(* CODESYS project Intecre_TwinSafeModels.library
   Author: Mark Lazarides
   Version: 0.5.0.3
   Description: Functional models of the TwinSAFE logic function blocks and TwinSAFE group, for trialling safety applications and their interaction with the standard PLC.
      
      0.4.2.0 - T_SafeFunctionBlockBase sets State to Run / Stop before Process; user FBs need no State logic.
      0.4.1.0 - corrects call issue with Example_UserFBs
      
      0.4.0.0 - Adds the eight channel (EL1918) and two channel (EL2912) terminal models.
      0.3.0.0 - Adds User FB examples, demonstrating extension.
   Title: Intecre.TwinSAFE.Models
   DefaultNamespace: Intecre.TwinSAFE.Models
   Placeholder: Intecre.TwinSAFE.Models
   Company: Intecre Ltd

Project tree, tasks and I/O mapping:
  libraries: Intecre.Utilities, * (Intecre Ltd); Tc2_Standard, * (Beckhoff Automation GmbH); Tc2_System, * (Beckhoff Automation GmbH); Tc3_Module, * (Beckhoff Automation GmbH); TcUnit, * (www.tcunit.org)
  Core/
    function F_NormaliseSafeInput [ST]
    function F_SafeInputValue [ST]
    function F_SafeResetTimeOk [ST]
    function block T_SafeConnection [ST]: FB_init, RunStateMachine, SetGroupReference, StateChanged
    function block T_SafeFunctionBlockBase [ST]: ClearDiagBit, ConfigurationOk, FB_init, Process, ReportRefusedConfiguration, SetDiagBit, SetGroupReference
    function block T_SafeGroup [ST]: ConnectionCount, FunctionBlockCount, GroupState, RaiseOnRefusedConfiguration, RegisterConnection, RegisterFunctionBlock, ScanMembers, StateChanged
    function block T_SafeInputPair [ST]
    function block T_SafeInputTerminal [ST]
    function block T_SafeInputTerminal8 [ST]
    function block T_SafeOutputTerminal [ST]
    function block T_SafeOutputTerminal2 [ST]
  DUTs/
    data type E_SafeConnectionError
    data type E_SafeConnectionState
    data type E_SafeEdmState
    data type E_SafeFbState
    data type E_SafeGroupDiag
    data type E_SafeGroupState
    data type E_SafeLatchState
    data type E_SafeMonState
    data type E_SafeMutingState
    data type E_SafeTonState
    data type E_SafeTwoHandState
    data type ST_SafeConnShutdownParameters
    data type ST_SafeEdmParameters
    data type ST_SafeEStopParameters
    data type ST_SafeLatchParameters
    data type ST_SafeLogicParameters
    data type ST_SafeMonParameters
    data type ST_SafeMutingParameters
    data type ST_SafeOpModeParameters
    data type ST_SafeTimerParameters
    data type ST_SafeTwoHandParameters
  Examples/
    Example_UserFbs/
      function block T_SafePulse_UserFB [CFC]: FB_init, Process
      function block T_SafeRTrig_UserFB [CFC]: FB_init, Process
    program PRG_EStopExample [ST]
    program PRG_EStopExample_CFC [CFC]
  FunctionBlocks/
    function block T_SafeAnd [ST]: ConfigurationOk, Process
    function block T_SafeConnShutdown [ST]: ConnShutdownState, FB_init, Process, StateChanged, UpdateDiscrepancyDiag
    function block T_SafeDecouple [ST]: Process
    function block T_SafeEdm [ST]: ConfigurationOk, Process, StateChanged
    function block T_SafeEStop [ST]: ConfigurationOk, EdmInputsOk, EdmInputsTrue, EdmResetOk, EStopState, Process, SetOutputsSafe, StartEdmResetMonitoring, StateChanged, UpdateDiscrepancyDiag
    function block T_SafeMon [ST]: ConfigurationOk, EdmInputsOk, EdmInputsTrue, EdmResetOk, MonState, Process, SetOutputsSafe, StartEdmResetMonitoring, StateChanged, UpdateDiscrepancyDiag
    function block T_SafeMuting [ST]: Actual, AddEvent, Advance, AnySensor, BuildSequence, ConfigurationOk, EdmInputsOk, EdmInputsTrue, EdmResetOk, IsMuting, MutingState, MutingStateFor, Process, SetOutputsSafe, StartEdmResetMonitoring, StateChanged, UpdateDiscrepancyDiag
    function block T_SafeOpMode [ST]: ConfigurationOk, Process, SetOutputs, StateChanged
    function block T_SafeOr [ST]: ConfigurationOk, Process
    function block T_SafeRs [ST]: ConfigurationOk, Process
    function block T_SafeSr [ST]: ConfigurationOk, Process
    function block T_SafeTof [ST]: ConfigurationOk, Process
    function block T_SafeTon [ST]: ConfigurationOk, Process
    function block T_SafeTwoHand [ST]: Process, SetHandDiscrepancyError, StateChanged, TwoHandState, UpdateDiscrepancyDiag
    function block T_SafeXor [ST]: Process
  Params/
    global variables SafeModelParams
  Project Information/
    function F_GetCompany [ST]
    function F_GetTitle [ST]
    function F_GetVersion [ST]
  Tests/
    User_FB_Tests/
      function block T_SafePulse_UserFB_Tests [ST]: Test_InnerBlocksJoinTheGroup, Test_PulseEndsWhenInputDrops, Test_PulseForDelayTimeWhileInputHeld, Test_StoppedGivesNoOutput
      function block T_SafePulse_UserFB_Tests_CFC [ST]: Test_InnerBlocksJoinTheGroup, Test_PulseEndsWhenInputDrops, Test_PulseForDelayTimeWhileInputHeld, Test_StoppedGivesNoOutput
      function block T_SafeRTrig_UserFB_Tests [ST]: Test_InnerBlocksJoinTheGroup, Test_StoppedGivesNoOutput, Test_TriggerForOneCycleOnRisingEdge
      function block T_SafeRTrig_UserFB_Tests_CFC [ST]: Test_InnerBlocksJoinTheGroup, Test_StoppedGivesNoOutput, Test_TriggerForOneCycleOnRisingEdge
    program PRG_TestRunner [ST]
    function block T_SafeAnd_Tests [ST]: Test_AllConnectedInputsTrueGivesRun, Test_OneConnectedInputIsRefused, Test_OneInputFalseGivesSafe, Test_RaiseOnRefusedConfigurationStopsHard, Test_StoppedGivesNoOutput, Test_UnconnectedInputsIgnoredAndMakeContactNegated
    function block T_SafeAnd_Tests_CFC [ST]: Test_AllConnectedInputsTrueGivesRun, Test_OneInputFalseGivesSafe, Test_StoppedGivesNoOutput, Test_UnconnectedInputsIgnoredAndMakeContactNegated
    function block T_SafeCfcTestSuite [ST]: FinishTest, StartTest
    function block T_SafeConnection_Tests [ST]: Test_ComErrorClearedByAcknowledge, Test_StartsUpToDataWhenGroupRuns
    function block T_SafeConnection_Tests_CFC [ST]: Test_ComErrorClearedByAcknowledge, Test_StartsUpToDataWhenGroupRuns
    function block T_SafeConnShutdown_Tests [ST]: Test_DeactivateShutsDownConnection
    function block T_SafeConnShutdown_Tests_CFC [ST]: Test_DeactivateShutsDownConnection
    function block T_SafeDecouple_Tests [ST]: Test_InputsLoopedToOutputsOnlyWhenRunning
    function block T_SafeDecouple_Tests_CFC [ST]: Test_InputsLoopedToOutputsOnlyWhenRunning
    function block T_SafeEdm_Tests [ST]: Test_NoErrorWhenFeedbackFollows, Test_SwitchOnTimeoutGivesError, Test_UnconnectedMon2IsRefused
    function block T_SafeEdm_Tests_CFC [ST]: Test_NoErrorWhenFeedbackFollows, Test_SwitchOnTimeoutGivesError
    function block T_SafeEStop_Tests [ST]: Test_DelayedOutput, Test_DiscrepancyErrorNeedsSafeInputsBeforeAck, Test_EdmErrorAtRestartAndAcknowledge, Test_EStopRequestSwitchesOutputsOffAndBlocksRestart, Test_MakeContactInputRequestsSafeStateOnOne, Test_OutputsOffWhenStopped, Test_ResetTimeOverSixtySecondsIsRefused, Test_RestartHeldBeforeEStopGivesEdmError, Test_StartupRequiresRestartSequence
    function block T_SafeEStop_Tests_CFC [ST]: Test_DelayedOutput, Test_DiscrepancyErrorNeedsSafeInputsBeforeAck, Test_EdmErrorAtRestartAndAcknowledge, Test_EStopRequestSwitchesOutputsOffAndBlocksRestart, Test_MakeContactInputRequestsSafeStateOnOne, Test_OutputsOffWhenStopped, Test_RestartHeldBeforeEStopGivesEdmError, Test_StartupRequiresRestartSequence
    function block T_SafeGroup_Tests [ST]: Test_ConnectionStartupAndComError, Test_FbErrorStopsGroupAndErrAckRecovers, Test_RefusesTheSixtyFifthConnection, Test_RegistersMoreThanSixtyFourBlocks, Test_RunsFunctionBlocksWithoutConnections, Test_StopWhenRunFalse
    function block T_SafeGroup_Tests_CFC [ST]: Test_ConnectionStartupAndComError, Test_FbErrorStopsGroupAndErrAckRecovers, Test_RunsFunctionBlocksWithoutConnections, Test_StopWhenRunFalse
    function block T_SafeInputPair_Tests [ST]: Test_BreakContactRequestsSafeStateOnZero, Test_DiscrepancyErrorAfterTimeoutAndResetAfterSafeInputs, Test_InactivePairNeverRequestsSafeState, Test_MakeContactRequestsSafeStateOnOne, Test_TwoChannelRequestsSafeStateIfEitherChannelLow
    function block T_SafeInputPair_Tests_CFC [ST]: Test_BreakContactRequestsSafeStateOnZero, Test_DiscrepancyErrorAfterTimeoutAndResetAfterSafeInputs, Test_InactivePairNeverRequestsSafeState, Test_MakeContactRequestsSafeStateOnOne, Test_TwoChannelRequestsSafeStateIfEitherChannelLow
    function block T_SafeInputTerminal8_Tests [ST]: Test_ComErrorForcesSafeInputsFalse, Test_RegistersAsConnection, Test_SafeInputsFalseBeforeData, Test_SafeInputsFollowChannelsInData
    function block T_SafeMon_Tests [ST]: Test_AutomaticRestartWhenGuardClosed, Test_EdmFaultWithoutManualRestartStaysSafe, Test_ManualFunctionTestRequiresGuardOpenedOnce, Test_NoMonInConnectedIsRefused, Test_ResetTimeNotMultipleOfTenIsRefused, Test_SecureInputBypassesGuard
    function block T_SafeMon_Tests_CFC [ST]: Test_AutomaticRestartWhenGuardClosed, Test_EdmFaultWithoutManualRestartStaysSafe, Test_ManualFunctionTestRequiresGuardOpenedOnce, Test_SecureInputBypassesGuard
    function block T_SafeMuting_Tests [ST]: Test_OssdBlockedWithoutMutingGivesSafe, Test_ResetTimeNotMultipleOfTenIsRefused, Test_SequenceViolationGivesError, Test_SequentialMutingKeepsOutputOn, Test_TwoSensorParallelSequence
    function block T_SafeMuting_Tests_CFC [ST]: Test_OssdBlockedWithoutMutingGivesSafe, Test_SequenceViolationGivesError, Test_SequentialMutingKeepsOutputOn, Test_TwoSensorParallelSequence
    function block T_SafeOpMode_Tests [ST]: Test_ConnectedRestartRequiresRestartSequence, Test_ExactlyOneInputSelectsOutput, Test_OneConnectedInputIsRefused, Test_SlowModeChangeGivesDiscrepancyError
    function block T_SafeOpMode_Tests_CFC [ST]: Test_ConnectedRestartRequiresRestartSequence, Test_ExactlyOneInputSelectsOutput, Test_SlowModeChangeGivesDiscrepancyError
    function block T_SafeOr_Tests [ST]: Test_AllFalseGivesSafe, Test_AnyConnectedInputTrueGivesRun, Test_OneConnectedInputIsRefused
    function block T_SafeOr_Tests_CFC [ST]: Test_AllFalseGivesSafe, Test_AnyConnectedInputTrueGivesRun
    function block T_SafeOutputTerminal2_Tests [ST]: Test_ChannelsFalseBeforeData, Test_ChannelsFollowSafeOutsInData, Test_ComErrorForcesChannelsFalse, Test_GroupNotRunningForcesChannelsFalse, Test_RegistersAsConnection
    function block T_SafeRs_Tests [ST]: Test_ResetDominantLatch, Test_UnconnectedSetIsRefused
    function block T_SafeRs_Tests_CFC [ST]: Test_ResetDominantLatch
    function block T_SafeSr_Tests [ST]: Test_SetDominantLatch, Test_UnconnectedResetIsRefused
    function block T_SafeSr_Tests_CFC [ST]: Test_SetDominantLatch
    function block T_SafeTof_Tests [ST]: Test_OutputDelayedOff, Test_UnconnectedInputIsRefused
    function block T_SafeTof_Tests_CFC [ST]: Test_OutputDelayedOff
    function block T_SafeTon_Tests [ST]: Test_OutputDelayedOn, Test_UnconnectedInputIsRefused
    function block T_SafeTon_Tests_CFC [ST]: Test_OutputDelayedOn
    function block T_SafeTwoHand_Tests [ST]: Test_BothHandsGiveOutputAndReleaseNeedsBothOff, Test_HandDiscrepancyTimeout, Test_SecondHandWithoutFirstGivesTwoHandError
    function block T_SafeTwoHand_Tests_CFC [ST]: Test_BothHandsGiveOutputAndReleaseNeedsBothOff, Test_HandDiscrepancyTimeout, Test_SecondHandWithoutFirstGivesTwoHandError
    function block T_SafeXor_Tests [ST]: Test_ConnectedPairsAreExclusiveOr
    function block T_SafeXor_Tests_CFC [ST]: Test_ConnectedPairsAreExclusiveOr
  Version/
    global variables Global_Version
*)

// DUTs/E_SafeConnectionError
// TwinSAFE connection error codes (low nibble of the connection Diag byte).
{attribute 'qualified_only'}
{attribute 'to_string'}
TYPE
E_SafeConnectionError :
(
    NoError := 0,
    InvalidCommand := 1,
    UnknownCommand := 2,
    InvalidConnectionId := 3,
    InvalidCrc := 4,
    WatchdogElapsed := 5,
    InvalidFsoeAddress := 6,
    InvalidData := 7,
    InvalidComParameterLength := 8,
    InvalidComParameters := 9,
    InvalidUserParameterLength := 10,
    InvalidUserParameters := 11,
    FsoeMasterReset := 12,
    SlaveModuleError := 13,
    OutputModuleError := 14,
    SlaveNotStarted := 15
) BYTE;
END_TYPE

// DUTs/E_SafeConnectionState
// TwinSAFE (FSoE) connection state codes.
{attribute 'qualified_only'}
{attribute 'to_string'}
TYPE
E_SafeConnectionState :
(
    Reset := 100,
    Session := 101,
    Connection := 102,
    Parameter := 103,
    Data := 104,
    Shutdown := 105,
    ShutdownDeactive := 106
) BYTE;
END_TYPE

// DUTs/E_SafeEdmState
// FB EDM state codes.
{attribute 'qualified_only'}
{attribute 'to_string'}
TYPE
E_SafeEdmState :
(
    Undefined := 0,
    Stop := 2,
    Error := 4,
    Reset := 5,
    MonOff := 14,
    MonOn := 15
) BYTE;
END_TYPE

// DUTs/E_SafeFbState
// TwinSAFE function block state codes shared by most FBs (Map State value).
// Error is also the state of a block whose configuration the TwinSAFE Safety Editor refuses (too few
// inputs connected, a required input unwired, an invalid EDM reset time): the block then sets Error,
// diagnostic bit 15 (16#8000), which no TwinSAFE FB uses, and stays in Error through every ErrAck.
// See T_SafeFunctionBlockBase.
{attribute 'qualified_only'}
{attribute 'to_string'}
TYPE
E_SafeFbState :
(
    Undefined := 0,
    Run := 1,
    Stop := 2,
    Safe := 3,
    Error := 4,
    Reset := 5,
    Start := 6,
    ErrorDelay := 7,
    DelayOut := 8
) BYTE;
END_TYPE

// DUTs/E_SafeGroupDiag
// TwinSAFE group diagnostic codes (EL/EJ6910).
{attribute 'qualified_only'}
{attribute 'to_string'}
TYPE
E_SafeGroupDiag :
(
    NoError := 0,
    FbError := 1,
    ComError := 2,
    ModuleError := 3,
    CmpError := 4,
    DeactivateError := 5,
    RestartError := 6
) BYTE;
END_TYPE

// DUTs/E_SafeGroupState
// TwinSAFE group state codes (EL/EJ6910).
{attribute 'qualified_only'}
{attribute 'to_string'}
TYPE
E_SafeGroupState :
(
    Undefined := 0,
    Run := 1,
    Stop := 2,
    Safe := 3,
    Error := 4,
    Reset := 5,
    Start := 6,
    StopError := 7,
    Deactive := 16,
    WaitComError := 17
) BYTE;
END_TYPE

// DUTs/E_SafeLatchState
// FB RS and FB SR state codes.
{attribute 'qualified_only'}
{attribute 'to_string'}
TYPE
E_SafeLatchState :
(
    Undefined := 0,
    Stop := 2,
    Safe := 3,
    Set := 9
) BYTE;
END_TYPE

// DUTs/E_SafeMonState
// FB MON state codes.
{attribute 'qualified_only'}
{attribute 'to_string'}
TYPE
E_SafeMonState :
(
    Undefined := 0,
    Run := 1,
    Stop := 2,
    Safe := 3,
    Error := 4,
    Reset := 5,
    Start := 6,
    ErrorDelay := 7,
    DelayOut := 8,
    FuncTest := 9
) BYTE;
END_TYPE

// DUTs/E_SafeMutingState
// FB MUTING state codes.
{attribute 'qualified_only'}
{attribute 'to_string'}
TYPE
E_SafeMutingState :
(
    Undefined := 0,
    Run := 1,
    Stop := 2,
    Safe := 3,
    Error := 4,
    Reset := 5,
    DelayOut := 8,
    Muting1 := 9,
    Muting2 := 10,
    Muting3 := 11,
    Muting4 := 12,
    Muting5 := 13,
    Muting6 := 14,
    Muting7 := 15,
    Muting8 := 16,
    Muting9 := 17
) BYTE;
END_TYPE

// DUTs/E_SafeTonState
// FB TON state codes.
{attribute 'qualified_only'}
{attribute 'to_string'}
TYPE
E_SafeTonState :
(
    Undefined := 0,
    Run := 1,
    Stop := 2,
    Safe := 3,
    DelayIn := 9
) BYTE;
END_TYPE

// DUTs/E_SafeTwoHandState
// FB TWOHAND state codes.
{attribute 'qualified_only'}
{attribute 'to_string'}
TYPE
E_SafeTwoHandState :
(
    Undefined := 0,
    Run := 1,
    Stop := 2,
    Safe := 3,
    Error := 4,
    Reset := 5,
    OneButton := 11,
    TwoButton := 12,
    Release := 13
) BYTE;
END_TYPE

// DUTs/ST_SafeConnShutdownParameters
// Parameters of FB CONNECTION SHUTDOWN.
TYPE
ST_SafeConnShutdownParameters :
STRUCT
    Deactivate1MakeContact : BOOL;
    Deactivate2MakeContact : BOOL;
    DiscrepancyTime : TIME;
    SafeInputsAfterDiscError : BOOL; // Safety Editor checkbox 'Safe Inputs after Disc Error', FALSE for a new block:
        // TRUE makes both channels of the pair that raised a discrepancy error return to the safe state together
        // before ErrAck can clear it
END_STRUCT
END_TYPE

// DUTs/ST_SafeEdmParameters
// Parameters of FB EDM.
TYPE
ST_SafeEdmParameters :
STRUCT
    Mon1MakeContact : BOOL;
    Mon2MakeContact : BOOL;
    SwitchOnTime : TIME; // Mon2 must become FALSE within this time of Mon1 rising. T#0S disables
    SwitchOffTime : TIME; // Mon2 must become TRUE within this time of Mon1 falling. T#0S disables
END_STRUCT
END_TYPE

// DUTs/ST_SafeEStopParameters
// Parameters of FB ESTOP (port and FB properties of the Safety Editor).
// Ports are active when connected; a pair is two channel when both ports are connected.
TYPE
ST_SafeEStopParameters :
STRUCT
    EStopIn1MakeContact : BOOL; // FALSE = break contact (0 requests the safe state); TRUE = make contact
    EStopIn2MakeContact : BOOL;
    EStopIn3MakeContact : BOOL;
    EStopIn4MakeContact : BOOL;
    EStopIn5MakeContact : BOOL;
    EStopIn6MakeContact : BOOL;
    EStopIn7MakeContact : BOOL;
    EStopIn8MakeContact : BOOL;
    DiscrepancyTime1 : TIME; // EStopIn1 / EStopIn2. T#0S = no discrepancy monitoring
    DiscrepancyTime2 : TIME; // EStopIn3 / EStopIn4
    DiscrepancyTime3 : TIME; // EStopIn5 / EStopIn6
    DiscrepancyTime4 : TIME; // EStopIn7 / EStopIn8
    DelayTime : TIME; // switch-off delay of EStopDelOut
    Edm1ResetTime : TIME; // EL6910: EDM1 must drop within this time of EStopOut switching on. T#0S disables
    Edm2ResetTime : TIME;
    SafeInputsAfterDiscError : BOOL; // Safety Editor checkbox, FALSE for a new block; the EL6910 always applies
        // 'Safe Inputs after Disc Error' to ESTOP whatever the box says (only the EL6900 honours it, and the editor
        // warns when it is TRUE under an EL6910), so the model ignores this value and always behaves as TRUE
END_STRUCT
END_TYPE

// DUTs/ST_SafeLatchParameters
// Parameters of FB RS and FB SR.
TYPE
ST_SafeLatchParameters :
STRUCT
    SetMakeContact : BOOL;
    ResetMakeContact : BOOL;
END_STRUCT
END_TYPE

// DUTs/ST_SafeLogicParameters
// Parameters of FB AND and FB OR. Inputs are active when connected.
TYPE
ST_SafeLogicParameters :
STRUCT
    In1MakeContact : BOOL; // TRUE = the input is negated before the logic operation
    In2MakeContact : BOOL;
    In3MakeContact : BOOL;
    In4MakeContact : BOOL;
    In5MakeContact : BOOL;
    In6MakeContact : BOOL;
    In7MakeContact : BOOL;
    In8MakeContact : BOOL;
END_STRUCT
END_TYPE

// DUTs/ST_SafeMonParameters
// Parameters of FB MON. Manual restart is active when the Restart port is connected.
TYPE
ST_SafeMonParameters :
STRUCT
    MonIn1MakeContact : BOOL;
    MonIn2MakeContact : BOOL;
    MonIn3MakeContact : BOOL;
    MonIn4MakeContact : BOOL;
    Secure1MakeContact : BOOL;
    Secure2MakeContact : BOOL;
    DiscrepancyTime1 : TIME; // MonIn1 / MonIn2
    DiscrepancyTime2 : TIME; // MonIn3 / MonIn4
    SecureDiscrepancyTime : TIME; // Secure1 / Secure2
    DelayTime : TIME; // switch-off delay of MonDelOut
    Edm1ResetTime : TIME;
    Edm2ResetTime : TIME;
    ManualFunctionTest : BOOL; // every connected MonIn pair must request the safe state once after start
    SafeInputsAfterDiscError : BOOL; // Safety Editor checkbox 'Safe Inputs after Disc Error', FALSE for a new block:
        // TRUE makes both channels of the pair that raised a discrepancy error return to the safe state together
        // before ErrAck can clear it
END_STRUCT
END_TYPE

// DUTs/ST_SafeMutingParameters
// Parameters of FB MUTING.
TYPE
ST_SafeMutingParameters :
STRUCT
    SequentialInputs : BOOL; // TRUE: single-channel muting sensors in sequence; FALSE: two two-channel sensors
    MutingIn1MakeContact : BOOL;
    MutingIn2MakeContact : BOOL;
    MutingIn3MakeContact : BOOL;
    MutingIn4MakeContact : BOOL;
    OSSDIn1MakeContact : BOOL;
    OSSDIn2MakeContact : BOOL;
    MutingDiscrepancyTime1 : TIME; // MutingIn1 / MutingIn2 (parallel mode)
    MutingDiscrepancyTime2 : TIME; // MutingIn3 / MutingIn4 (parallel mode)
    OssdDiscrepancyTime : TIME; // OSSDIn1 / OSSDIn2
    FilterTime : TIME; // debounce of the muting inputs (max 500 ms)
    MaxMutingTime : TIME; // max duration of a muting sequence (max 10 min). T#0S disables
    DelayTime : TIME; // switch-off delay of MuteDelOut (max 30 s)
    Edm1ResetTime : TIME;
    Edm2ResetTime : TIME;
    BackwardsMode : BOOL; // EL6910: sequence may also run from the last sensor to the first
    OssdCheckOptional : BOOL; // EL6910: protective device is not part of the sequence check
    SafeInputsAfterDiscError : BOOL; // Safety Editor checkbox 'Safe Inputs after Disc Error', FALSE for a new block:
        // TRUE makes both channels of the pair that raised a discrepancy error return to the safe state together
        // before ErrAck can clear it
END_STRUCT
END_TYPE

// DUTs/ST_SafeOpModeParameters
// Parameters of FB OPMODE. Manual restart is active when the Restart port is connected.
TYPE
ST_SafeOpModeParameters :
STRUCT
    DiscrepancyTime : TIME; // max time during a mode change with none or several inputs set. T#0S disables
END_STRUCT
END_TYPE

// DUTs/ST_SafeTimerParameters
// Parameters of FB TON and FB TOF.
TYPE
ST_SafeTimerParameters :
STRUCT
    MakeContact : BOOL;
    DelayTime : TIME;
END_STRUCT
END_TYPE

// DUTs/ST_SafeTwoHandParameters
// Parameters of FB TWOHAND.
TYPE
ST_SafeTwoHandParameters :
STRUCT
    Twohand1MakeContact : BOOL;
    Twohand2MakeContact : BOOL;
    Twohand3MakeContact : BOOL;
    Twohand4MakeContact : BOOL;
    DiscrepancyTime1 : TIME; // Twohand1 / Twohand2
    DiscrepancyTime2 : TIME; // Twohand3 / Twohand4
    HandDiscrepancyTime : TIME; // max time between actuation of the two hands (max 2500 ms). T#0S disables
    SafeInputsAfterDiscError : BOOL; // Safety Editor checkbox 'Safe Inputs after Disc Error', FALSE for a new block:
        // TRUE makes both channels of the pair that raised a discrepancy error return to the safe state together
        // before ErrAck can clear it
END_STRUCT
END_TYPE

// Params/SafeModelParams
// Library parameters of Intecre.TwinSAFE.Models: the project-wide defaults, set per project in the
// Library Manager's parameter view without rebuilding the library. A parameter list must be constant,
// so the run-time switch lives on T_SafeGroup (RaiseOnRefusedConfiguration), initialised from here.
{attribute 'qualified_only'}
VAR_GLOBAL CONSTANT
    // Default of T_SafeGroup.RaiseOnRefusedConfiguration for every group. TRUE: a block of the group whose
    // configuration the TwinSAFE Safety Editor refuses (see T_SafeFunctionBlockBase) raises
    // RTSEXCPT_IO_CONFIG_ERROR with F_RaiseException after it has reported Error, so the controller stops
    // on the first cycle unless the call is in a __TRY block. FALSE: the block only reports Error,
    // State = Error and diagnostic bit 15, and logs the fault once.
    RAISE_ON_REFUSED_CONFIGURATION : BOOL := FALSE;
END_VAR

// Version/Global_Version
{attribute 'TcGenerated'}
{attribute 'no-analysis'}
{attribute 'linkalways'}
// This function has been automatically generated from the project information.
VAR_GLOBAL CONSTANT
	{attribute 'const_non_replaced'}
	stLibVersion_Intecre_TwinSAFE_Models : ST_LibVersion := (iMajor := 0, iMinor := 5, iBuild := 0, iRevision := 3, nFlags := 0, sVersion := '0.5.0.3');
END_VAR

// Core/F_NormaliseSafeInput
// Applies the port configuration to a raw input value.
// Result TRUE means "not requesting the safe state" (the released / healthy condition).
// An unconnected (inactive) port never requests the safe state.
FUNCTION F_NormaliseSafeInput : BOOL
VAR_INPUT
    active : BOOL; // port is connected
    makeContact : BOOL; // FALSE = break contact (0 requests the safe state), TRUE = make contact (signal negated)
    value : BOOL;
END_VAR

IF NOT active THEN
    F_NormaliseSafeInput := TRUE;
    RETURN;
END_IF

F_NormaliseSafeInput := value XOR makeContact;

END_FUNCTION

// Core/F_SafeInputValue
// Applies the port configuration to a raw input value for ports that assert a function
// (Set, Reset, TonIn, OrIn, muting sensors ...). An unconnected port reads FALSE.
FUNCTION F_SafeInputValue : BOOL
VAR_INPUT
    active : BOOL;
    makeContact : BOOL;
    value : BOOL;
END_VAR

IF NOT active THEN
    F_SafeInputValue := FALSE;
    RETURN;
END_IF

F_SafeInputValue := value XOR makeContact;

END_FUNCTION

// Core/F_SafeResetTimeOk
// TRUE when an EDM 'Reset Time' parameter is one the Safety Editor accepts: 0 ms (off) or a multiple
// of 10 ms, and at most 60000 ms. The editor reports "'Reset Time' parameter ... has to be 0 ms or a
// multiple of 10 ms and maximal 60000 ms" otherwise.
FUNCTION F_SafeResetTimeOk : BOOL
VAR_INPUT
    resetTime : TIME;
END_VAR
VAR CONSTANT
    MAX_RESET_TIME : TIME := T#60S;
END_VAR

IF resetTime > MAX_RESET_TIME THEN
    RETURN;
END_IF

F_SafeResetTimeOk := (TIME_TO_UDINT(resetTime) MOD 10 = 0);

END_FUNCTION

// Core/T_SafeConnection
// Simulated TwinSAFE (FSoE) connection between the logic and a safe I/O terminal or another logic.
// Belongs to a group from construction:  conn : T_SafeConnection(group := safetyGroup);
// Starts up through Reset -> Session -> Connection -> Parameter -> Data once the group runs.
// Communication errors are injected with InjectComError and cleared by the group ErrAck
// (plus ComErrAck when ComErrAckActive is set).
FUNCTION_BLOCK T_SafeConnection
VAR_INPUT
    ComErrAck : BOOL; // connection specific acknowledgement (EL6910 option ComErrAckActive)
    LocalShutdown : BOOL; // shutdown requested by FB CONNECTION SHUTDOWN (set through its reference)
    PartnerShutdown : BOOL; // simulates a shutdown command received from the FSoE partner
    InjectComError : BOOL; // rising edge simulates an FSoE communication error
    InjectErrorCode : E_SafeConnectionError := E_SafeConnectionError.WatchdogElapsed;
    StartupTime : TIME := T#300MS; // simulated time from Reset to Data
    ComErrAckActive : BOOL; // connection needs its own ComErrAck in addition to the group ErrAck
END_VAR
VAR_OUTPUT
    ComError : BOOL;
    InStartup : BOOL;
    InDataState : BOOL;
    OutputsEnabled : BOOL; // in the Data state with the group in RUN: the only time a safe output terminal passes its SafeOut values (a group in STOP or ERROR switches every output of the group off)
    IsShutdown : BOOL;
    State : BYTE; // connection state code 100..106
    Diag : BYTE; // connection diagnostic byte
END_VAR
VAR
    _group : REFERENCE TO T_SafeGroup;
    _state : E_SafeConnectionState := E_SafeConnectionState.Reset;
    _prevState : E_SafeConnectionState;
    _errorCode : E_SafeConnectionError;
    _groupAcknowledged : BOOL;
    _comErrAcked : BOOL;
    _errAckPrev : BOOL;
    _comErrAckPrev : BOOL;
    _injectPrev : BOOL;
    _startupTimer : TON;
END_VAR

IF NOT __ISVALIDREF(_group) THEN
    RETURN; // not (yet) assigned to a group: stays in its initial (fail-safe) state
END_IF

IF _group.ErrAck AND NOT _errAckPrev THEN
    _groupAcknowledged := TRUE;
END_IF

_errAckPrev := _group.ErrAck;

IF ComErrAck AND NOT _comErrAckPrev THEN
    _comErrAcked := TRUE;
END_IF

_comErrAckPrev := ComErrAck;

IF InjectComError AND NOT _injectPrev THEN
    ComError           := TRUE;
    _errorCode         := InjectErrorCode;
    _groupAcknowledged := FALSE;
    _comErrAcked       := FALSE;
    _state             := E_SafeConnectionState.Reset;
END_IF

_injectPrev := InjectComError;

// A communication error is cleared once the group (and if required the connection) has acknowledged.
IF ComError AND _groupAcknowledged AND (NOT ComErrAckActive OR _comErrAcked) THEN
    ComError           := FALSE;
    _errorCode         := E_SafeConnectionError.NoError;
    _groupAcknowledged := FALSE;
    _comErrAcked       := FALSE;
END_IF

RunStateMachine();

InStartup := NOT ComError
                 AND (_state = E_SafeConnectionState.Reset
                 OR _state = E_SafeConnectionState.Session
                 OR _state = E_SafeConnectionState.Connection
                 OR _state = E_SafeConnectionState.Parameter);

InDataState := (_state = E_SafeConnectionState.Data);
OutputsEnabled := InDataState AND _group.InRun;
IsShutdown  := (_state = E_SafeConnectionState.Shutdown) OR (_state = E_SafeConnectionState.ShutdownDeactive);
State       := TO_BYTE(_state);
Diag        := TO_BYTE(_errorCode);

IF InStartup THEN
    Diag := Diag OR 16#40;
END_IF

IF ComError THEN
    Diag := Diag OR 16#10;
END_IF

METHOD FB_init : BOOL
VAR_INPUT
    bInitRetains : BOOL;
    bInCopyCode : BOOL;
    group : REFERENCE TO T_SafeGroup; // the TwinSAFE group this connection is assigned to
END_VAR
SetGroupReference(
    bInCopyCode := bInCopyCode,
    group := group
);
END_METHOD

METHOD PRIVATE RunStateMachine
VAR
    stepTime : TIME;
END_VAR
stepTime := UDINT_TO_TIME(TIME_TO_UDINT(StartupTime) / 3);

CASE _state OF
    E_SafeConnectionState.Reset:
        IF StateChanged() THEN
            _startupTimer(IN := FALSE, PT := stepTime);
        END_IF

        IF _group.Run AND NOT ComError THEN
            _state := E_SafeConnectionState.Session;
        END_IF

    E_SafeConnectionState.Session:
        IF StateChanged() THEN
            _startupTimer(IN := FALSE, PT := stepTime);
        END_IF

        _startupTimer(IN := TRUE, PT := stepTime);

        IF _startupTimer.Q THEN
            _state := E_SafeConnectionState.Connection;
        END_IF

    E_SafeConnectionState.Connection:
        IF StateChanged() THEN
            _startupTimer(IN := FALSE, PT := stepTime);
        END_IF

        _startupTimer(IN := TRUE, PT := stepTime);

        IF _startupTimer.Q THEN
            _state := E_SafeConnectionState.Parameter;
        END_IF

    E_SafeConnectionState.Parameter:
        IF StateChanged() THEN
            _startupTimer(IN := FALSE, PT := stepTime);
        END_IF

        _startupTimer(IN := TRUE, PT := stepTime);

        IF _startupTimer.Q THEN
            _state := E_SafeConnectionState.Data;
        END_IF

    E_SafeConnectionState.Data:
        StateChanged();

        IF LocalShutdown THEN
            _state := E_SafeConnectionState.ShutdownDeactive;
        ELSIF PartnerShutdown THEN
            _state := E_SafeConnectionState.Shutdown;
        END_IF

    E_SafeConnectionState.Shutdown:
        StateChanged();

        IF NOT PartnerShutdown THEN
            _state := E_SafeConnectionState.Reset;
        END_IF

    E_SafeConnectionState.ShutdownDeactive:
        StateChanged();

        IF NOT LocalShutdown THEN
            _state := E_SafeConnectionState.Reset;
        END_IF
END_CASE
END_METHOD

// Assigns the connection to a TwinSAFE group and registers it there. Called by FB_init; call it
// yourself from the FB_init of a composite (user) block to pass its group on to a connection it
// contains, which was declared with the composite's own _group before that reference was valid.
// Registering twice with the same group is harmless. Returns TRUE when the group was valid.
METHOD PUBLIC SetGroupReference : BOOL
VAR_INPUT
    bInCopyCode : BOOL;
    group : REFERENCE TO T_SafeGroup; // the TwinSAFE group this connection is assigned to
END_VAR
IF NOT __ISVALIDREF(group) THEN
    RETURN;
END_IF

_group REF= group;

IF NOT bInCopyCode THEN
    group.RegisterConnection(THIS^);
END_IF

SetGroupReference := TRUE;
END_METHOD

METHOD PRIVATE StateChanged : BOOL
IF _prevState = _state THEN
    RETURN;
END_IF

_prevState   := _state;
StateChanged := TRUE;
END_METHOD

END_FUNCTION_BLOCK

// Core/T_SafeGroup
// Model of a TwinSAFE group (EL/EJ6910 semantics).
// Function blocks and connections join the group at construction (FB_init group reference) and the
// group reads their outputs, so nothing needs wiring beyond the standard PLC signals.
// Call the group before its members each cycle. Declare the group before its members.
// RaiseOnRefusedConfiguration (default SafeModelParams.RAISE_ON_REFUSED_CONFIGURATION) makes a member
// whose configuration the Safety Editor refuses stop the controller with F_RaiseException after it has
// reported Error; see T_SafeFunctionBlockBase.
FUNCTION_BLOCK T_SafeGroup
VAR_INPUT
    Run : BOOL := TRUE; // Run/Stop. Link to a standard PLC variable.
    ErrAck : BOOL; // Error acknowledge (FALSE -> TRUE -> FALSE). Link to a standard PLC variable.
    ModuleFault : BOOL; // error input from another module (e.g. EK1960)
END_VAR
VAR_OUTPUT
    ComErr : BOOL; // communication error in at least one connection
    FbErr : BOOL; // at least one FB is in the ERROR state
    OutErr : BOOL; // not used (local outputs only exist on KL6904)
    OtherErr : BOOL; // ModuleFault
    ComStartup : BOOL; // at least one connection is starting up
    FbDeactive : BOOL; // group deactivated by customising (not modelled, always FALSE)
    FbRun : BOOL; // all FBs are in the RUN state
    InRun : BOOL; // the group is in the RUN state (FbRun of the members)
    State : BYTE; // group state code (Map State)
    Diag : BYTE; // group diagnostic code (Map Diag)
    RegistrationRefused : BOOL; // a block or connection could not join because the group is full (MAX_FUNCTION_BLOCKS, MAX_CONNECTIONS): the model is then incomplete, never expected in use
END_VAR
VAR CONSTANT
    MAX_FUNCTION_BLOCKS : UINT := 256;
    MAX_CONNECTIONS : UINT := 64;
END_VAR
VAR
    _functionBlocks : ARRAY[1..MAX_FUNCTION_BLOCKS] OF POINTER TO T_SafeFunctionBlockBase;
    _functionBlockCount : UINT;
    _connections : ARRAY[1..MAX_CONNECTIONS] OF POINTER TO T_SafeConnection;
    _connectionCount : UINT;
    _state : E_SafeGroupState := E_SafeGroupState.Stop;
    _prevState : E_SafeGroupState;
    _errAckPrev : BOOL;
    _errAckFallingEdge : BOOL;
    _anyFbError : BOOL;
    _allFbsRunning : BOOL;
    _anyComError : BOOL;
    _anyComStartup : BOOL;
    _anyError : BOOL;
    _raiseOnRefusedConfiguration : BOOL := SafeModelParams.RAISE_ON_REFUSED_CONFIGURATION;
END_VAR

_errAckFallingEdge := NOT ErrAck AND _errAckPrev;
_errAckPrev        := ErrAck;
ScanMembers();
_anyError := _anyFbError OR _anyComError OR ModuleFault;

CASE _state OF
    E_SafeGroupState.Undefined,
    E_SafeGroupState.Stop:
        StateChanged();

        IF _anyError THEN
            _state := E_SafeGroupState.StopError;
        ELSIF Run THEN
            _state := SEL(_anyComStartup, E_SafeGroupState.Run, E_SafeGroupState.Start);
        END_IF

    E_SafeGroupState.StopError:
        StateChanged();

        IF Run THEN
            _state := E_SafeGroupState.Error;
        ELSIF NOT _anyError THEN
            _state := E_SafeGroupState.Stop;
        END_IF

    E_SafeGroupState.Start:
        StateChanged();

        IF _anyError THEN
            _state := E_SafeGroupState.Error;
        ELSIF NOT Run THEN
            _state := E_SafeGroupState.Stop;
        ELSIF NOT _anyComStartup THEN
            _state := E_SafeGroupState.Run;
        END_IF

    E_SafeGroupState.Run:
        StateChanged();

        IF _anyError THEN
            _state := E_SafeGroupState.Error;
        ELSIF NOT Run THEN
            _state := E_SafeGroupState.Stop;
        ELSIF _anyComStartup THEN
            _state := E_SafeGroupState.Start;
        END_IF

    E_SafeGroupState.Error:
        StateChanged();

        IF NOT Run THEN
            _state := E_SafeGroupState.StopError;
        ELSIF ErrAck AND NOT _anyError THEN
            _state := E_SafeGroupState.Reset;
        END_IF

    E_SafeGroupState.Reset:
        StateChanged();

        IF _anyError THEN
            _state := E_SafeGroupState.Error;
        ELSIF _errAckFallingEdge THEN
            IF NOT Run THEN
                _state := E_SafeGroupState.Stop;
            ELSIF _anyComStartup THEN
                _state := E_SafeGroupState.Start;
            ELSE
                _state := E_SafeGroupState.Run;
            END_IF
        END_IF

ELSE
    _state := E_SafeGroupState.Stop;
END_CASE

ComErr     := _anyComError;
FbErr      := _anyFbError;
OutErr     := FALSE;
OtherErr   := ModuleFault;
ComStartup := _anyComStartup;
FbDeactive := FALSE;
FbRun      := _allFbsRunning;
InRun      := (_state = E_SafeGroupState.Run);
State      := TO_BYTE(_state);

IF _anyFbError THEN
    Diag := TO_BYTE(E_SafeGroupDiag.FbError);
ELSIF _anyComError THEN
    Diag := TO_BYTE(E_SafeGroupDiag.ComError);
ELSIF ModuleFault THEN
    Diag := TO_BYTE(E_SafeGroupDiag.ModuleError);
ELSE
    Diag := TO_BYTE(E_SafeGroupDiag.NoError);
END_IF

PROPERTY ConnectionCount : UINT
GET
ConnectionCount := _connectionCount;
END_GET
END_PROPERTY

PROPERTY FunctionBlockCount : UINT
GET
FunctionBlockCount := _functionBlockCount;
END_GET
END_PROPERTY

PROPERTY GroupState : E_SafeGroupState
GET
GroupState := _state;
END_GET
END_PROPERTY

// TRUE: a member whose configuration the TwinSAFE Safety Editor refuses raises RTSEXCPT_IO_CONFIG_ERROR
// (F_RaiseException) after reporting Error, so the controller stops unless the call is in a __TRY block.
// Starts at SafeModelParams.RAISE_ON_REFUSED_CONFIGURATION; set it per group from project code or a test.
PROPERTY RaiseOnRefusedConfiguration : BOOL
GET
RaiseOnRefusedConfiguration := _raiseOnRefusedConfiguration;
END_GET
SET
_raiseOnRefusedConfiguration := RaiseOnRefusedConfiguration;
END_SET
END_PROPERTY

// Called by T_SafeConnection.FB_init. Not part of the public interface.
METHOD INTERNAL RegisterConnection
VAR_INPUT
    connection : REFERENCE TO T_SafeConnection;
END_VAR
VAR
    i : UINT;
END_VAR
FOR i := 1 TO _connectionCount DO
    IF _connections[i] = ADR(connection) THEN
        RETURN;
    END_IF
END_FOR

IF _connectionCount >= MAX_CONNECTIONS THEN
    RegistrationRefused := TRUE;
    RETURN;
END_IF

_connectionCount               := _connectionCount + 1;
_connections[_connectionCount] := ADR(connection);
END_METHOD

// Called by T_SafeFunctionBlockBase.FB_init. Not part of the public interface.
METHOD INTERNAL RegisterFunctionBlock
VAR_INPUT
    functionBlock : REFERENCE TO T_SafeFunctionBlockBase;
END_VAR
VAR
    i : UINT;
END_VAR
FOR i := 1 TO _functionBlockCount DO
    IF _functionBlocks[i] = ADR(functionBlock) THEN
        RETURN;
    END_IF
END_FOR

IF _functionBlockCount >= MAX_FUNCTION_BLOCKS THEN
    RegistrationRefused := TRUE;
    RETURN;
END_IF

_functionBlockCount                  := _functionBlockCount + 1;
_functionBlocks[_functionBlockCount] := ADR(functionBlock);
END_METHOD

// Reads the outputs of the registered function blocks and connections.
METHOD PRIVATE ScanMembers
VAR
    i : UINT;
END_VAR
_anyFbError    := FALSE;
_allFbsRunning := (_functionBlockCount > 0);

FOR i := 1 TO _functionBlockCount DO
    _anyFbError    := _anyFbError OR _functionBlocks[i]^.Error;
    _allFbsRunning := _allFbsRunning AND _functionBlocks[i]^.IsRunning;
END_FOR

_anyComError   := FALSE;
_anyComStartup := FALSE;

FOR i := 1 TO _connectionCount DO
    _anyComError   := _anyComError OR _connections[i]^.ComError;
    _anyComStartup := _anyComStartup OR _connections[i]^.InStartup;
END_FOR
END_METHOD

METHOD PRIVATE StateChanged : BOOL
IF _prevState = _state THEN
    RETURN;
END_IF

_prevState   := _state;
StateChanged := TRUE;
END_METHOD

END_FUNCTION_BLOCK

// Core/T_SafeFunctionBlockBase
// Common behaviour of every modelled TwinSAFE function block.
// A block belongs to a TwinSAFE group from construction: declare it as
//     eStop : T_SafeEStop(group := safetyGroup);
// It registers with the group, takes FbRun (group in RUN) and ErrAck from it, and the group
// reads its Error and IsRunning outputs. Declare the group before its members.
// Derived classes implement Process(). Before Process() the base sets State to Run while the group
// runs and to Stop otherwise, so a block built only from other blocks needs no State logic; a block
// with states of its own overwrites State in Process(), and writes Error and Diag when it has them.
//
// Configuration check. The Safety Editor refuses some wirings and parameter values at project verify
// (an AND with one input, an SR with Reset unwired, an EDM reset time that is not a multiple of 10 ms).
// A block with such a rule overrides ConfigurationOk() and writes the editor's message to
// _configurationFault when the rule is broken. The base then runs the block as a stopped block (outputs
// at their safe value), reports Error with State = Error and diagnostic bit 15 (16#8000, a bit no
// TwinSAFE FB uses), logs the fault once through the Intecre.Utilities logger with the instance name in
// front (taken from the private T_NamedBase member _log; the project has to set LogConfig.LogLevel to
// Error or lower, as the logger is silent by default), and keeps the error through every ErrAck: a
// configuration error cannot be acknowledged away, only rewired.
// With the group's RaiseOnRefusedConfiguration TRUE (default SafeModelParams.RAISE_ON_REFUSED_CONFIGURATION,
// a library parameter) the base also raises RTSEXCPT_IO_CONFIG_ERROR with F_RaiseException after
// reporting, so a simulation stops hard on the first cycle unless the call sits in a __TRY block
// (a __CATCH on 4026 receives a TwinCAT code, not RTSEXCPT_IO_CONFIG_ERROR; check Error and Diag).
FUNCTION_BLOCK ABSTRACT T_SafeFunctionBlockBase
VAR_OUTPUT
    Error : BOOL; // FB Error output
    State : BYTE; // FB state code (Map State)
    Diag : WORD; // FB diagnostic bits (Map Diag)
    IsRunning : BOOL; // FB in the RUN state
END_VAR
VAR CONSTANT
    CONFIGURATION_REFUSED_DIAG_BIT : INT := 15; // Diag bit set while the Safety Editor would refuse the configuration
END_VAR
VAR
    _group : REFERENCE TO T_SafeGroup;
    _fbRun : BOOL; // group in RUN
    _errAck : BOOL; // group error acknowledge
    _errAckPrev : BOOL;
    _errAckRisingEdge : BOOL;
    _errAckFallingEdge : BOOL;
    _configurationRefused : BOOL; // ConfigurationOk() returned FALSE this cycle
    _configurationFault : T_MaxString; // the editor's message for the broken rule, written by ConfigurationOk()
    _configurationLogged : BOOL; // the fault has been logged (once per instance)
    _log : T_NamedBase; // supplies the instance path for the log line; its InstanceName ends in ._log, which ReportRefusedConfiguration trims
END_VAR

IF __ISVALIDREF(_group) THEN
    _fbRun  := _group.InRun;
    _errAck := _group.ErrAck;
ELSE
    // not (yet) in a group: behaves as a stopped block until SetGroupReference is called
    _fbRun  := FALSE;
    _errAck := FALSE;
END_IF

_configurationRefused := NOT ConfigurationOk();

IF _configurationRefused THEN
    // the Safety Editor refuses this wiring or parameter set: the block runs as a stopped block, so its
    // outputs take their safe value, and the error reported below is not acknowledged
    _fbRun  := FALSE;
    _errAck := FALSE;
END_IF

_errAckRisingEdge  := _errAck AND NOT _errAckPrev;
_errAckFallingEdge := NOT _errAck AND _errAckPrev;
_errAckPrev        := _errAck;
// default state: Run while the group runs, else Stop. Blocks with states of their own overwrite it in
// Process(). Error and Diag are not reset here: they latch until ErrAck in TwinSAFE, so only the block
// that raised them clears them.
State := TO_BYTE(SEL(_fbRun, E_SafeFbState.Stop, E_SafeFbState.Run));
Process();

IF _configurationRefused THEN
    Error := TRUE;
    State := TO_BYTE(E_SafeFbState.Error);
    SetDiagBit(CONFIGURATION_REFUSED_DIAG_BIT);
END_IF

IsRunning := (State = TO_BYTE(E_SafeFbState.Run));

IF _configurationRefused THEN
    ReportRefusedConfiguration();
END_IF

METHOD PROTECTED ClearDiagBit
VAR_INPUT
    bitIndex : INT;
END_VAR
Diag := Diag AND NOT SHL(WORD#1, bitIndex);
END_METHOD

// TRUE when the block is wired and parameterised as the TwinSAFE Safety Editor accepts it. A block
// with a rule overrides this method; when the rule is broken it writes the editor's own message to
// _configurationFault and returns FALSE. The base then reports the block in Error (see the header).
METHOD PROTECTED ConfigurationOk : BOOL
ConfigurationOk := TRUE;
END_METHOD

METHOD FB_init : BOOL
VAR_INPUT
    bInitRetains : BOOL;
    bInCopyCode : BOOL;
    group : REFERENCE TO T_SafeGroup; // the TwinSAFE group this block belongs to
END_VAR
SetGroupReference(
    bInCopyCode := bInCopyCode,
    group := group
);
END_METHOD

METHOD PROTECTED ABSTRACT Process
END_METHOD

// Logs the refused configuration once per instance as '<instance>: <block type>: <editor's rule> (...)',
// the instance being _log.InstanceName minus its own '._log' segment, then stops the controller with
// RTSEXCPT_IO_CONFIG_ERROR when the group's RaiseOnRefusedConfiguration asks for it (a block without a
// group follows the library parameter). Called after Error, State and Diag have been written, so a
// __CATCH sees the block already in Error. The logger is Intecre.Utilities' F_LogError, which is silent
// until the project sets LogConfig.LogLevel.
METHOD PRIVATE ReportRefusedConfiguration
VAR
    instance : T_MaxString;
    raise : BOOL;
END_VAR
VAR CONSTANT
    MEMBER_SUFFIX : STRING := '._log';
END_VAR
IF NOT _configurationLogged THEN
    _configurationLogged := TRUE;
    instance := _log.InstanceName;

    IF RIGHT(instance, LEN(MEMBER_SUFFIX)) = MEMBER_SUFFIX THEN
        instance := LEFT(instance, LEN(instance) - LEN(MEMBER_SUFFIX));
    END_IF

    F_LogError(CONCAT(CONCAT(instance, ': '), CONCAT(_configurationFault, ' (the TwinSAFE Safety Editor refuses this configuration)')));
END_IF

IF __ISVALIDREF(_group) THEN
    raise := _group.RaiseOnRefusedConfiguration;
ELSE
    raise := SafeModelParams.RAISE_ON_REFUSED_CONFIGURATION;
END_IF

IF raise THEN
    F_RaiseException(TO_UDINT(__SYSTEM.ExceptionCode.RTSEXCPT_IO_CONFIG_ERROR));
END_IF
END_METHOD

METHOD PROTECTED SetDiagBit
VAR_INPUT
    bitIndex : INT;
END_VAR
Diag := Diag OR SHL(WORD#1, bitIndex);
END_METHOD

// Assigns the block to a TwinSAFE group and registers it there. Called by FB_init; call it
// yourself from the FB_init of a composite (user) block to pass its group on to the blocks it
// contains, which were declared with the composite's own _group before that reference was valid.
// Registering twice with the same group is harmless. Returns TRUE when the group was valid.
METHOD PUBLIC SetGroupReference : BOOL
VAR_INPUT
    bInCopyCode : BOOL;
    group : REFERENCE TO T_SafeGroup; // the TwinSAFE group this block belongs to
END_VAR
IF NOT __ISVALIDREF(group) THEN
    RETURN;
END_IF

_group REF= group;

IF NOT bInCopyCode THEN
    group.RegisterFunctionBlock(THIS^);
END_IF

SetGroupReference := TRUE;
END_METHOD

END_FUNCTION_BLOCK

// FunctionBlocks/T_SafeEStop
// Model of the TwinSAFE FB ESTOP.
// Up to eight emergency stop inputs in four pairs, immediate and delayed outputs,
// two feedback loops (EDM) and a manual restart requiring a 0 -> 1 -> 0 sequence on Restart.
// Ports are active when connected.
// The Safety Editor refuses an EDM reset time that is not 0 ms, a multiple of 10 ms and at most 60000 ms:
// the model then reports Error with diagnostic bit 15 instead of running (see T_SafeFunctionBlockBase).
{attribute 'reflection'}
FUNCTION_BLOCK T_SafeEStop EXTENDS T_SafeFunctionBlockBase
VAR_INPUT
    Restart : BOOL; // may be a standard PLC signal
    EDM1 : BOOL; // feedback loop of EStopOut (may be a standard PLC signal)
    EDM2 : BOOL; // feedback loop of EStopDelOut (may be a standard PLC signal)
    EStopIn1 : BOOL;
    EStopIn2 : BOOL;
    EStopIn3 : BOOL;
    EStopIn4 : BOOL;
    EStopIn5 : BOOL;
    EStopIn6 : BOOL;
    EStopIn7 : BOOL;
    EStopIn8 : BOOL;
    Parameters : ST_SafeEStopParameters;
END_VAR
VAR_OUTPUT
    EStopOut : BOOL; // switches off immediately
    EStopDelOut : BOOL; // switches off after DelayTime
END_VAR
VAR
    {attribute 'is_connected' := 'Restart'}
    _restartConnected : BOOL;
    {attribute 'is_connected' := 'EDM1'}
    _eDM1Connected : BOOL;
    {attribute 'is_connected' := 'EDM2'}
    _eDM2Connected : BOOL;
    {attribute 'is_connected' := 'EStopIn1'}
    _eStopIn1Connected : BOOL;
    {attribute 'is_connected' := 'EStopIn2'}
    _eStopIn2Connected : BOOL;
    {attribute 'is_connected' := 'EStopIn3'}
    _eStopIn3Connected : BOOL;
    {attribute 'is_connected' := 'EStopIn4'}
    _eStopIn4Connected : BOOL;
    {attribute 'is_connected' := 'EStopIn5'}
    _eStopIn5Connected : BOOL;
    {attribute 'is_connected' := 'EStopIn6'}
    _eStopIn6Connected : BOOL;
    {attribute 'is_connected' := 'EStopIn7'}
    _eStopIn7Connected : BOOL;
    {attribute 'is_connected' := 'EStopIn8'}
    _eStopIn8Connected : BOOL;
    _pairs : ARRAY[1..4] OF T_SafeInputPair;
    _state : E_SafeFbState := E_SafeFbState.Stop;
    _prevState : E_SafeFbState;
    _restartPrev : BOOL;
    _delayTimer : TON;
    _edmResetTimer1 : TON;
    _edmResetTimer2 : TON;
    _edm1Dropped : BOOL;
    _edm2Dropped : BOOL;
END_VAR

SUPER^();

// The EDM reset times must be 0 ms or a multiple of 10 ms up to 60000 ms (Safety Editor: "'Reset Time' parameter ... has to be 0 ms or a multiple of 10 ms and maximal 60000 ms").
METHOD PROTECTED ConfigurationOk : BOOL
IF NOT F_SafeResetTimeOk(Parameters.Edm1ResetTime) THEN
    _configurationFault := 'T_SafeEStop: $'Reset Time$' parameter of EDM1 of ESTOP has to be 0 ms or a multiple of 10 ms and maximal 60000 ms';
    RETURN;
ELSIF NOT F_SafeResetTimeOk(Parameters.Edm2ResetTime) THEN
    _configurationFault := 'T_SafeEStop: $'Reset Time$' parameter of EDM2 of ESTOP has to be 0 ms or a multiple of 10 ms and maximal 60000 ms';
    RETURN;
END_IF

ConfigurationOk := TRUE;
END_METHOD

// Checks the EDM inputs at restart and records diagnostic bits 4/5 on failure.
METHOD PRIVATE EdmInputsOk : BOOL
EdmInputsOk := TRUE;

IF _eDM1Connected AND NOT EDM1 THEN
    SetDiagBit(4);
    EdmInputsOk := FALSE;
END_IF

IF _eDM2Connected AND NOT EDM2 THEN
    SetDiagBit(5);
    EdmInputsOk := FALSE;
END_IF
END_METHOD

// TRUE when every connected EDM input reads 1 (contactors released).
METHOD PRIVATE EdmInputsTrue : BOOL
EdmInputsTrue := (NOT _eDM1Connected OR EDM1) AND (NOT _eDM2Connected OR EDM2);
END_METHOD

// EL6910 extension: after the outputs switch on, each connected EDM input must drop to FALSE
// within its Reset Time. Returns FALSE (and sets diagnostic bits 4/5) on timeout.
METHOD PRIVATE EdmResetOk : BOOL
EdmResetOk := TRUE;

IF _eDM1Connected AND Parameters.Edm1ResetTime > T#0S THEN
    IF NOT EDM1 THEN
        _edm1Dropped := TRUE;
    END_IF

    _edmResetTimer1(IN := NOT _edm1Dropped, PT := Parameters.Edm1ResetTime);

    IF _edmResetTimer1.Q THEN
        SetDiagBit(4);
        EdmResetOk := FALSE;
    END_IF
END_IF

IF _eDM2Connected AND Parameters.Edm2ResetTime > T#0S THEN
    IF NOT EDM2 THEN
        _edm2Dropped := TRUE;
    END_IF

    _edmResetTimer2(IN := NOT _edm2Dropped, PT := Parameters.Edm2ResetTime);

    IF _edmResetTimer2.Q THEN
        SetDiagBit(5);
        EdmResetOk := FALSE;
    END_IF
END_IF
END_METHOD

PROPERTY EStopState : E_SafeFbState
GET
EStopState := _state;
END_GET
END_PROPERTY

METHOD PROTECTED Process
VAR
    i : USINT;
    acknowledge : BOOL;
    safeRequested : BOOL;
    discError : BOOL;
    restartFalling : BOOL;
    operating : BOOL;
    stateBefore : E_SafeFbState;
    passes : USINT;
END_VAR
acknowledge := (_state = E_SafeFbState.Error) AND _errAck;
_pairs[1](
    In1 := EStopIn1,
    In2 := EStopIn2,
    Active1 := _eStopIn1Connected,
    Active2 := _eStopIn2Connected,
    MakeContact1 := Parameters.EStopIn1MakeContact,
    MakeContact2 := Parameters.EStopIn2MakeContact,
    DiscrepancyTime := Parameters.DiscrepancyTime1,
    Monitor := _fbRun,
    SafeInputsAfterDiscError := TRUE, // the EL6910 always applies it to ESTOP, whatever the parameter says
    Acknowledge := acknowledge
);

_pairs[2](
    In1 := EStopIn3,
    In2 := EStopIn4,
    Active1 := _eStopIn3Connected,
    Active2 := _eStopIn4Connected,
    MakeContact1 := Parameters.EStopIn3MakeContact,
    MakeContact2 := Parameters.EStopIn4MakeContact,
    DiscrepancyTime := Parameters.DiscrepancyTime2,
    Monitor := _fbRun,
    SafeInputsAfterDiscError := TRUE, // the EL6910 always applies it to ESTOP, whatever the parameter says
    Acknowledge := acknowledge
);

_pairs[3](
    In1 := EStopIn5,
    In2 := EStopIn6,
    Active1 := _eStopIn5Connected,
    Active2 := _eStopIn6Connected,
    MakeContact1 := Parameters.EStopIn5MakeContact,
    MakeContact2 := Parameters.EStopIn6MakeContact,
    DiscrepancyTime := Parameters.DiscrepancyTime3,
    Monitor := _fbRun,
    SafeInputsAfterDiscError := TRUE, // the EL6910 always applies it to ESTOP, whatever the parameter says
    Acknowledge := acknowledge
);

_pairs[4](
    In1 := EStopIn7,
    In2 := EStopIn8,
    Active1 := _eStopIn7Connected,
    Active2 := _eStopIn8Connected,
    MakeContact1 := Parameters.EStopIn7MakeContact,
    MakeContact2 := Parameters.EStopIn8MakeContact,
    DiscrepancyTime := Parameters.DiscrepancyTime4,
    Monitor := _fbRun,
    SafeInputsAfterDiscError := TRUE, // the EL6910 always applies it to ESTOP, whatever the parameter says
    Acknowledge := acknowledge
);

FOR i := 1 TO 4 DO
    safeRequested := safeRequested OR _pairs[i].SafeStateRequested;
    discError     := discError OR _pairs[i].DiscrepancyError;
END_FOR

restartFalling := NOT Restart AND _restartPrev;
_restartPrev   := Restart;

IF NOT _fbRun AND _state <> E_SafeFbState.Error AND _state <> E_SafeFbState.Reset THEN
    _state := E_SafeFbState.Stop;
END_IF

// A discrepancy error is detected in every operating state
operating := (_state = E_SafeFbState.Safe)
                 OR (_state = E_SafeFbState.Start)
                 OR (_state = E_SafeFbState.Run)
                 OR (_state = E_SafeFbState.DelayOut);

IF discError AND operating THEN
    UpdateDiscrepancyDiag();
    _state := E_SafeFbState.Error;
END_IF

passes := 0;

REPEAT
    stateBefore := _state;

    CASE _state OF
        E_SafeFbState.Stop:
            IF StateChanged() THEN
                SetOutputsSafe();
                Error := FALSE;
                Diag  := 0;
            END_IF

            IF _fbRun THEN
                _state := E_SafeFbState.Safe;
            END_IF

        E_SafeFbState.Safe:
            IF StateChanged() THEN
                SetOutputsSafe();
            END_IF

            // A TRUE restart signal triggers the EDM check immediately (see restart behaviour sample 3)
            IF Restart THEN
                IF NOT EdmInputsOk() THEN
                    _state := E_SafeFbState.Error;
                ELSIF NOT safeRequested THEN
                    _state := E_SafeFbState.Start;
                END_IF
            END_IF

        E_SafeFbState.Start:
            IF StateChanged() THEN
                SetOutputsSafe();
            END_IF

            IF safeRequested THEN
                _state := E_SafeFbState.Safe;
            ELSIF restartFalling THEN
                IF EdmInputsOk() THEN
                    _state := E_SafeFbState.Run;
                ELSE
                    _state := E_SafeFbState.Error;
                END_IF
            END_IF

        E_SafeFbState.Run:
            IF StateChanged() THEN
                EStopOut    := TRUE;
                EStopDelOut := TRUE;
                StartEdmResetMonitoring();
            END_IF

            IF NOT EdmResetOk() THEN
                _state := E_SafeFbState.Error;
            ELSIF safeRequested THEN
                IF Parameters.DelayTime > T#0S THEN
                    _state := E_SafeFbState.DelayOut;
                ELSE
                    _state := E_SafeFbState.Safe;
                END_IF
            END_IF

        E_SafeFbState.DelayOut:
            IF StateChanged() THEN
                EStopOut    := FALSE;
                EStopDelOut := TRUE;
                _delayTimer(IN := FALSE, PT := Parameters.DelayTime);
            END_IF

            _delayTimer(IN := TRUE, PT := Parameters.DelayTime);

            IF _delayTimer.Q THEN
                _state := E_SafeFbState.Safe;
            END_IF

        E_SafeFbState.Error:
            IF StateChanged() THEN
                SetOutputsSafe();
                Error := TRUE;
            END_IF

            UpdateDiscrepancyDiag();

            IF _errAck AND NOT discError THEN
                _state := E_SafeFbState.Reset;
            END_IF

        E_SafeFbState.Reset:
            IF StateChanged() THEN
                SetOutputsSafe();
                Error := FALSE;
                Diag  := 0;
            END_IF

            IF _errAckFallingEdge THEN
                _state := SEL(_fbRun, E_SafeFbState.Stop, E_SafeFbState.Safe);
            END_IF
    END_CASE

    passes := passes + 1;
UNTIL (stateBefore = _state) OR (passes >= 3)
END_REPEAT

State := TO_BYTE(_state);
END_METHOD

METHOD PRIVATE SetOutputsSafe
EStopOut    := FALSE;
EStopDelOut := FALSE;
END_METHOD

METHOD PRIVATE StartEdmResetMonitoring
_edm1Dropped := FALSE;
_edm2Dropped := FALSE;
_edmResetTimer1(IN := FALSE, PT := Parameters.Edm1ResetTime);
_edmResetTimer2(IN := FALSE, PT := Parameters.Edm2ResetTime);
END_METHOD

METHOD PRIVATE StateChanged : BOOL
IF _prevState = _state THEN
    RETURN;
END_IF

_prevState   := _state;
StateChanged := TRUE;
END_METHOD

// Mirrors the discrepancy state of every pair into the diagnostic bits.
METHOD PRIVATE UpdateDiscrepancyDiag
VAR
    i : USINT;
END_VAR
FOR i := 1 TO 4 DO
    IF _pairs[i].DiscrepancyError THEN
        SetDiagBit(i - 1);

        IF _pairs[i].AwaitingSafeInputs THEN
            SetDiagBit(i + 7);
        ELSE
            ClearDiagBit(i + 7);
        END_IF
    END_IF
END_FOR
END_METHOD

END_FUNCTION_BLOCK

// Core/T_SafeInputPair
// Evaluates a one- or two-channel FB input pair with optional discrepancy monitoring,
// exactly as the TwinSAFE FBs treat their paired inputs (EStopIn1/2, MonIn1/2, Twohand1/2 ...).
// Internal helper used by the modelled FBs.
FUNCTION_BLOCK T_SafeInputPair
VAR_INPUT
    In1 : BOOL;
    In2 : BOOL;
    Active1 : BOOL; // channel 1 port is connected
    Active2 : BOOL; // channel 2 port is connected
    MakeContact1 : BOOL;
    MakeContact2 : BOOL;
    DiscrepancyTime : TIME; // T#0S = two channel without discrepancy monitoring
    Monitor : BOOL; // discrepancy monitoring runs only while TRUE (FB executed by a running group)
    SafeInputsAfterDiscError : BOOL; // both channels must be safe together before a discrepancy error can be acknowledged
    Acknowledge : BOOL; // clear a discrepancy error this cycle if permitted
END_VAR
VAR_OUTPUT
    Channel1 : BOOL; // normalised: TRUE = not requesting the safe state
    Channel2 : BOOL;
    IsActive : BOOL;
    IsTwoChannel : BOOL;
    AllTrue : BOOL; // all active channels TRUE (TRUE when inactive)
    AllFalse : BOOL; // all active channels FALSE (FALSE when inactive)
    SafeStateRequested : BOOL;
    DiscrepancyError : BOOL;
    AwaitingSafeInputs : BOOL;
END_VAR
VAR
    _discrepancyTimer : TON;
END_VAR

Channel1     := F_NormaliseSafeInput(Active1, MakeContact1, In1);
Channel2     := F_NormaliseSafeInput(Active2, MakeContact2, In2);
IsActive     := Active1 OR Active2;
IsTwoChannel := Active1 AND Active2;

IF Monitor AND IsTwoChannel AND DiscrepancyTime > T#0S THEN
    _discrepancyTimer(IN := (Channel1 <> Channel2), PT := DiscrepancyTime);

    IF _discrepancyTimer.Q AND NOT DiscrepancyError THEN
        DiscrepancyError   := TRUE;
        AwaitingSafeInputs := SafeInputsAfterDiscError;
    END_IF
ELSE
    _discrepancyTimer(IN := FALSE, PT := DiscrepancyTime);
END_IF

IF AwaitingSafeInputs AND NOT Channel1 AND NOT Channel2 THEN
    AwaitingSafeInputs := FALSE;
END_IF

IF Acknowledge AND DiscrepancyError AND NOT AwaitingSafeInputs THEN
    DiscrepancyError := FALSE;
    _discrepancyTimer(IN := FALSE, PT := DiscrepancyTime);
END_IF

AllTrue            := Channel1 AND Channel2;
AllFalse           := IsActive AND (NOT Active1 OR NOT Channel1) AND (NOT Active2 OR NOT Channel2);
SafeStateRequested := NOT AllTrue;

END_FUNCTION_BLOCK

// Core/T_SafeInputTerminal
// Model of a four channel safe input terminal (EL1904): a TwinSAFE connection with four channels.
// Declare it in its group:  inputTerminal : T_SafeInputTerminal(group := safetyGroup);
// Channel1..4 are the simulated field signals; SafeIn1..4 are what the TwinSAFE logic sees:
// forced FALSE (fail-safe) unless the connection is in the Data state.
FUNCTION_BLOCK T_SafeInputTerminal EXTENDS T_SafeConnection
VAR_INPUT
    Channel1 : BOOL;
    Channel2 : BOOL;
    Channel3 : BOOL;
    Channel4 : BOOL;
END_VAR
VAR_OUTPUT
    SafeIn1 : BOOL;
    SafeIn2 : BOOL;
    SafeIn3 : BOOL;
    SafeIn4 : BOOL;
END_VAR

SUPER^();
SafeIn1 := Channel1 AND InDataState;
SafeIn2 := Channel2 AND InDataState;
SafeIn3 := Channel3 AND InDataState;
SafeIn4 := Channel4 AND InDataState;

END_FUNCTION_BLOCK

// Core/T_SafeInputTerminal8
// Model of an eight channel safe input terminal (EL1918): a TwinSAFE connection with eight channels.
// Declare it in its group:  inputTerminal : T_SafeInputTerminal8(group := safetyGroup);
// Channel1..8 are the simulated field signals; SafeIn1..8 are what the TwinSAFE logic sees:
// forced FALSE (fail-safe) unless the connection is in the Data state.
FUNCTION_BLOCK T_SafeInputTerminal8 EXTENDS T_SafeConnection
VAR_INPUT
    Channel1 : BOOL;
    Channel2 : BOOL;
    Channel3 : BOOL;
    Channel4 : BOOL;
    Channel5 : BOOL;
    Channel6 : BOOL;
    Channel7 : BOOL;
    Channel8 : BOOL;
END_VAR
VAR_OUTPUT
    SafeIn1 : BOOL;
    SafeIn2 : BOOL;
    SafeIn3 : BOOL;
    SafeIn4 : BOOL;
    SafeIn5 : BOOL;
    SafeIn6 : BOOL;
    SafeIn7 : BOOL;
    SafeIn8 : BOOL;
END_VAR

SUPER^();
SafeIn1 := Channel1 AND InDataState;
SafeIn2 := Channel2 AND InDataState;
SafeIn3 := Channel3 AND InDataState;
SafeIn4 := Channel4 AND InDataState;
SafeIn5 := Channel5 AND InDataState;
SafeIn6 := Channel6 AND InDataState;
SafeIn7 := Channel7 AND InDataState;
SafeIn8 := Channel8 AND InDataState;

END_FUNCTION_BLOCK

// Core/T_SafeOutputTerminal
// Model of a four channel safe output terminal (EL2904): a TwinSAFE connection with four channels.
// Declare it in its group:  outputTerminal : T_SafeOutputTerminal(group := safetyGroup);
// SafeOut1..4 are wired from FB outputs; Channel1..4 are the simulated field outputs,
// forced FALSE (fail-safe) unless the connection is in the Data state and the group is in RUN (OutputsEnabled).
FUNCTION_BLOCK T_SafeOutputTerminal EXTENDS T_SafeConnection
VAR_INPUT
    SafeOut1 : BOOL;
    SafeOut2 : BOOL;
    SafeOut3 : BOOL;
    SafeOut4 : BOOL;
END_VAR
VAR_OUTPUT
    Channel1 : BOOL;
    Channel2 : BOOL;
    Channel3 : BOOL;
    Channel4 : BOOL;
END_VAR

SUPER^();
Channel1 := SafeOut1 AND OutputsEnabled;
Channel2 := SafeOut2 AND OutputsEnabled;
Channel3 := SafeOut3 AND OutputsEnabled;
Channel4 := SafeOut4 AND OutputsEnabled;

END_FUNCTION_BLOCK

// Core/T_SafeOutputTerminal2
// Model of a two channel safe output terminal (EL2912): a TwinSAFE connection with two channels.
// Declare it in its group:  outputTerminal : T_SafeOutputTerminal2(group := safetyGroup);
// SafeOut1..2 are wired from FB outputs; Channel1..2 are the simulated field outputs,
// forced FALSE (fail-safe) unless the connection is in the Data state and the group is in RUN (OutputsEnabled).
FUNCTION_BLOCK T_SafeOutputTerminal2 EXTENDS T_SafeConnection
VAR_INPUT
    SafeOut1 : BOOL;
    SafeOut2 : BOOL;
END_VAR
VAR_OUTPUT
    Channel1 : BOOL;
    Channel2 : BOOL;
END_VAR

SUPER^();
Channel1 := SafeOut1 AND OutputsEnabled;
Channel2 := SafeOut2 AND OutputsEnabled;

END_FUNCTION_BLOCK

// Examples/Example_UserFbs/T_SafePulse_UserFB
FUNCTION_BLOCK T_SafePulse_UserFB EXTENDS T_SafeFunctionBlockBase
VAR_INPUT
	TonIn1 : BOOL;
	Parameters : ST_SafeTimerParameters;
END_VAR
VAR_OUTPUT
	TonOut : BOOL;
END_VAR
VAR
	safeTon : T_SafeTon(_group);
	safeAnd : T_SafeAnd(_group);
END_VAR

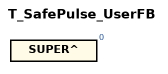
SUPER^();

METHOD FB_init : BOOL
VAR_INPUT
	bInitRetains	: BOOL;
	bInCopyCode	: BOOL;
	group	: REFERENCE TO T_SafeGroup;
END_VAR
safeAnd.SetGroupReference(bInCopyCode := bInCopyCode, group := group);
safeTon.SetGroupReference(bInCopyCode := bInCopyCode, group := group);
END_METHOD

METHOD PROTECTED Process
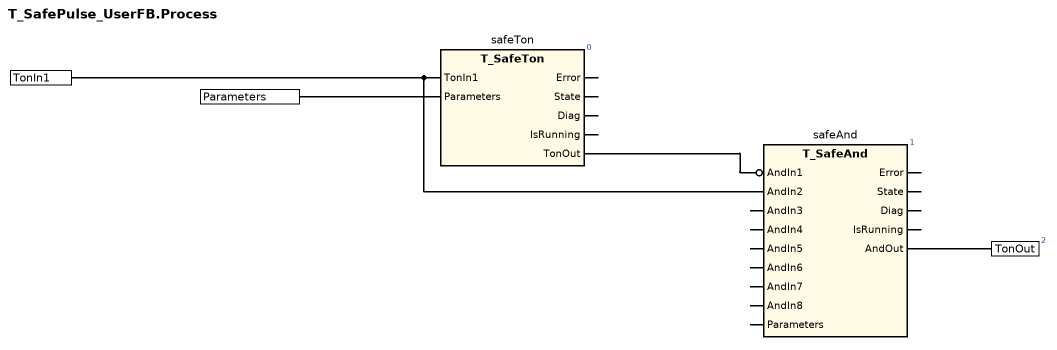
safeTon(TonIn1 := TonIn1, Parameters := Parameters); // T_SafeTon
safeAnd(AndIn1 := NOT safeTon.TonOut, AndIn2 := TonIn1); // T_SafeAnd
TonOut := safeAnd.AndOut;
END_METHOD

END_FUNCTION_BLOCK

// FunctionBlocks/T_SafeTon
// Model of the TwinSAFE FB TON (switch-on delay).
// The Safety Editor refuses a TON with TonIn1 unconnected: the model then reports Error with diagnostic
// bit 15 instead of running (see T_SafeFunctionBlockBase).
{attribute 'reflection'}
FUNCTION_BLOCK T_SafeTon EXTENDS T_SafeFunctionBlockBase
VAR_INPUT
    TonIn1 : BOOL;
    Parameters : ST_SafeTimerParameters;
END_VAR
VAR_OUTPUT
    TonOut : BOOL;
END_VAR
VAR
    {attribute 'is_connected' := 'TonIn1'}
    _tonIn1Connected : BOOL;
    _state : E_SafeTonState := E_SafeTonState.Stop;
    _timer : TON;
END_VAR

SUPER^();

// TonIn1 must be connected (Safety Editor: "Inport TonIn1 of TON must be connected").
METHOD PROTECTED ConfigurationOk : BOOL
IF NOT _tonIn1Connected THEN
    _configurationFault := 'T_SafeTon: Inport TonIn1 of TON must be connected';
    RETURN;
END_IF

ConfigurationOk := TRUE;
END_METHOD

METHOD PROTECTED Process
VAR
    inputActive : BOOL;
END_VAR
inputActive := _fbRun AND F_SafeInputValue(_tonIn1Connected, Parameters.MakeContact, TonIn1);
_timer(IN := inputActive, PT := Parameters.DelayTime);

IF NOT _fbRun THEN
    _state := E_SafeTonState.Stop;
ELSIF NOT inputActive THEN
    _state := E_SafeTonState.Safe;
ELSIF _timer.Q THEN
    _state := E_SafeTonState.Run;
ELSE
    _state := E_SafeTonState.DelayIn;
END_IF

TonOut := (_state = E_SafeTonState.Run);
Error  := FALSE;
Diag   := 0;
State  := TO_BYTE(_state);
END_METHOD

END_FUNCTION_BLOCK

// FunctionBlocks/T_SafeAnd
// Model of the TwinSAFE FB AND. Connected inputs are active; AndIn1 may be a standard PLC signal.
// The Safety Editor refuses an AND with fewer than two AndIn ports connected: the model then reports
// Error with diagnostic bit 15 instead of running (see T_SafeFunctionBlockBase).
{attribute 'reflection'}
FUNCTION_BLOCK T_SafeAnd EXTENDS T_SafeFunctionBlockBase
VAR_INPUT
    AndIn1 : BOOL;
    AndIn2 : BOOL;
    AndIn3 : BOOL;
    AndIn4 : BOOL;
    AndIn5 : BOOL;
    AndIn6 : BOOL;
    AndIn7 : BOOL;
    AndIn8 : BOOL;
    Parameters : ST_SafeLogicParameters;
END_VAR
VAR_OUTPUT
    AndOut : BOOL;
END_VAR
VAR
    {attribute 'is_connected' := 'AndIn1'}
    _andIn1Connected : BOOL;
    {attribute 'is_connected' := 'AndIn2'}
    _andIn2Connected : BOOL;
    {attribute 'is_connected' := 'AndIn3'}
    _andIn3Connected : BOOL;
    {attribute 'is_connected' := 'AndIn4'}
    _andIn4Connected : BOOL;
    {attribute 'is_connected' := 'AndIn5'}
    _andIn5Connected : BOOL;
    {attribute 'is_connected' := 'AndIn6'}
    _andIn6Connected : BOOL;
    {attribute 'is_connected' := 'AndIn7'}
    _andIn7Connected : BOOL;
    {attribute 'is_connected' := 'AndIn8'}
    _andIn8Connected : BOOL;
    _state : E_SafeFbState := E_SafeFbState.Stop;
END_VAR

SUPER^();

// At least two AndIn ports must be connected (Safety Editor: "AND does not have at least 2 input ports active and connected").
METHOD PROTECTED ConfigurationOk : BOOL
VAR
    connectedInputs : USINT;
END_VAR
connectedInputs := BOOL_TO_USINT(_andIn1Connected)
    + BOOL_TO_USINT(_andIn2Connected)
    + BOOL_TO_USINT(_andIn3Connected)
    + BOOL_TO_USINT(_andIn4Connected)
    + BOOL_TO_USINT(_andIn5Connected)
    + BOOL_TO_USINT(_andIn6Connected)
    + BOOL_TO_USINT(_andIn7Connected)
    + BOOL_TO_USINT(_andIn8Connected);

IF connectedInputs < 2 THEN
    _configurationFault := 'T_SafeAnd: AND does not have at least 2 input ports active and connected';
    RETURN;
END_IF

ConfigurationOk := TRUE;
END_METHOD

METHOD PROTECTED Process
VAR
    result : BOOL;
END_VAR
result := TRUE;
result := result AND F_NormaliseSafeInput(_andIn1Connected, Parameters.In1MakeContact, AndIn1);
result := result AND F_NormaliseSafeInput(_andIn2Connected, Parameters.In2MakeContact, AndIn2);
result := result AND F_NormaliseSafeInput(_andIn3Connected, Parameters.In3MakeContact, AndIn3);
result := result AND F_NormaliseSafeInput(_andIn4Connected, Parameters.In4MakeContact, AndIn4);
result := result AND F_NormaliseSafeInput(_andIn5Connected, Parameters.In5MakeContact, AndIn5);
result := result AND F_NormaliseSafeInput(_andIn6Connected, Parameters.In6MakeContact, AndIn6);
result := result AND F_NormaliseSafeInput(_andIn7Connected, Parameters.In7MakeContact, AndIn7);
result := result AND F_NormaliseSafeInput(_andIn8Connected, Parameters.In8MakeContact, AndIn8);

IF NOT _fbRun THEN
    _state := E_SafeFbState.Stop;
ELSIF result THEN
    _state := E_SafeFbState.Run;
ELSE
    _state := E_SafeFbState.Safe;
END_IF

AndOut := (_state = E_SafeFbState.Run);
Error  := FALSE;
Diag   := 0;
State  := TO_BYTE(_state);
END_METHOD

END_FUNCTION_BLOCK

// Examples/Example_UserFbs/T_SafeRTrig_UserFB
FUNCTION_BLOCK T_SafeRTrig_UserFB EXTENDS T_SafeFunctionBlockBase
VAR_INPUT
	Signal : BOOL;
END_VAR
VAR_OUTPUT
	Trigger : BOOL;
END_VAR
VAR
	safeRs : T_SafeRs(_group);
	safeAnd : T_SafeAnd(_group);
END_VAR

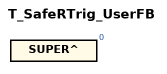
SUPER^();

METHOD FB_init : BOOL
VAR_INPUT
	bInitRetains	: BOOL;
	bInCopyCode	: BOOL;
	group	: REFERENCE TO T_SafeGroup;
END_VAR
safeRs.SetGroupReference(bInCopyCode := bInCopyCode, group := group);
safeAnd.SetGroupReference(bInCopyCode := bInCopyCode, group := group);
END_METHOD

METHOD PROTECTED Process
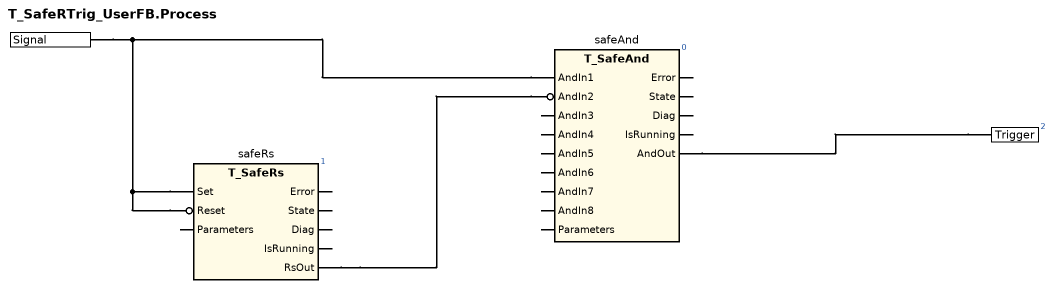
safeAnd(AndIn1 := Signal, AndIn2 := NOT safeRs.RsOut); // T_SafeAnd
safeRs(Set := Signal, Reset := NOT Signal); // T_SafeRs
Trigger := safeAnd.AndOut;
END_METHOD

END_FUNCTION_BLOCK

// FunctionBlocks/T_SafeRs
// Model of the TwinSAFE FB RS (reset dominant latch).
// The Safety Editor refuses an RS with Set or Reset unconnected: the model then reports Error with
// diagnostic bit 15 instead of running (see T_SafeFunctionBlockBase).
{attribute 'reflection'}
FUNCTION_BLOCK T_SafeRs EXTENDS T_SafeFunctionBlockBase
VAR_INPUT
    Set : BOOL;
    Reset : BOOL;
    Parameters : ST_SafeLatchParameters;
END_VAR
VAR_OUTPUT
    RsOut : BOOL;
END_VAR
VAR
    {attribute 'is_connected' := 'Set'}
    _setConnected : BOOL;
    {attribute 'is_connected' := 'Reset'}
    _resetConnected : BOOL;
    _state : E_SafeLatchState := E_SafeLatchState.Stop;
END_VAR

SUPER^();

// Set and Reset must both be connected (Safety Editor: "Inport Set of RS must be connected").
METHOD PROTECTED ConfigurationOk : BOOL
IF NOT _setConnected THEN
    _configurationFault := 'T_SafeRs: Inport Set of RS must be connected';
    RETURN;
ELSIF NOT _resetConnected THEN
    _configurationFault := 'T_SafeRs: Inport Reset of RS must be connected';
    RETURN;
END_IF

ConfigurationOk := TRUE;
END_METHOD

METHOD PROTECTED Process
VAR
    setActive : BOOL;
    resetActive : BOOL;
END_VAR
setActive   := F_SafeInputValue(_setConnected, Parameters.SetMakeContact, Set);
resetActive := F_SafeInputValue(_resetConnected, Parameters.ResetMakeContact, Reset);

IF NOT _fbRun THEN
    _state := E_SafeLatchState.Stop;
ELSE
    IF _state = E_SafeLatchState.Stop THEN
        _state := E_SafeLatchState.Safe;
    END_IF

    IF resetActive THEN
        _state := E_SafeLatchState.Safe;
    ELSIF setActive THEN
        _state := E_SafeLatchState.Set;
    END_IF
END_IF

RsOut := (_state = E_SafeLatchState.Set);
Error := FALSE;
Diag  := 0;
State := TO_BYTE(_state);
END_METHOD

END_FUNCTION_BLOCK

// Examples/PRG_EStopExample
// Worked example: a two-channel emergency stop with contactor feedback, wired the way a
// TwinSAFE project links it, plus the standard PLC signals (Run, ErrAck, Restart).
// The blocks join the group at declaration; call the group before its members.
// Toggle the "field" variables online to trial the behaviour and watch the State / Diag outputs.
PROGRAM PRG_EStopExample
VAR
    // --- simulated field devices (real hardware in a TwinSAFE system)
    eStopChannel1 : BOOL := TRUE; // NC contact, TRUE = not pressed
    eStopChannel2 : BOOL := TRUE;

    // --- standard PLC interface to the TwinSAFE group (linked to standard variables)
    safetyRun : BOOL := TRUE;
    safetyErrAck : BOOL;
    restartButton : BOOL; // 0 -> 1 -> 0 to restart

    // --- TwinSAFE model: the group, then its members (parameters as in the Safety Editor property grid)
    group : T_SafeGroup;
    inputTerminal : T_SafeInputTerminal(group := group); // EL1904
    outputTerminal : T_SafeOutputTerminal(group := group); // EL2904
    eStop : T_SafeEStop(group := group) := (Parameters := (DiscrepancyTime1 := T#500MS, DelayTime := T#1S));

    // --- simulated contactors: pull in 50 ms after the safe output energises; EDM1 = NOT pulled in
    contactorPullIn : TON;
END_VAR

// TwinSAFE group: standard PLC signals in; it reads its members' states itself
group(Run := safetyRun, ErrAck := safetyErrAck);

// Field -> safe input terminal (EL1904)
inputTerminal(Channel1 := eStopChannel1, Channel2 := eStopChannel2);

// FB ESTOP wired as in the safety project: EStopIn1/2 two channel, EDM1 and Restart from standard signals
eStop(
    Restart := restartButton,
    EDM1 := NOT contactorPullIn.Q,
    EStopIn1 := inputTerminal.SafeIn1,
    EStopIn2 := inputTerminal.SafeIn2
);

// Safe outputs -> output terminal (EL2904) -> field
outputTerminal(SafeOut1 := eStop.EStopOut, SafeOut2 := eStop.EStopDelOut);

// Simulated contactors follow the field output
contactorPullIn(IN := outputTerminal.Channel1, PT := T#50MS);

END_PROGRAM

// Examples/PRG_EStopExample_CFC
// Worked example: a two-channel emergency stop with contactor feedback, wired the way a
// TwinSAFE project links it, plus the standard PLC signals (Run, ErrAck, Restart).
// The blocks join the group at declaration; call the group before its members.
// CFC twin of PRG_EStopExample: the same wiring as a diagram.
// Toggle the "field" variables online to trial the behaviour and watch the State / Diag outputs.
PROGRAM PRG_EStopExample_CFC
VAR
    // --- simulated field devices (real hardware in a TwinSAFE system)
    eStopChannel1 : BOOL := TRUE; // NC contact, TRUE = not pressed
    eStopChannel2 : BOOL := TRUE;

    // --- standard PLC interface to the TwinSAFE group (linked to standard variables)
    safetyRun : BOOL := TRUE;
    safetyErrAck : BOOL;
    restartButton : BOOL; // 0 -> 1 -> 0 to restart

    // --- TwinSAFE model: the group, then its members (parameters as in the Safety Editor property grid)
    group : T_SafeGroup;
    inputTerminal : T_SafeInputTerminal(group := group); // EL1904
    outputTerminal : T_SafeOutputTerminal(group := group); // EL2904
    eStop : T_SafeEStop(group := group) := (Parameters := (DiscrepancyTime1 := T#500MS, DelayTime := T#1S));

    // --- simulated contactors: pull in 50 ms after the safe output energises; EDM1 = NOT pulled in
    contactorPullIn : TON;
END_VAR

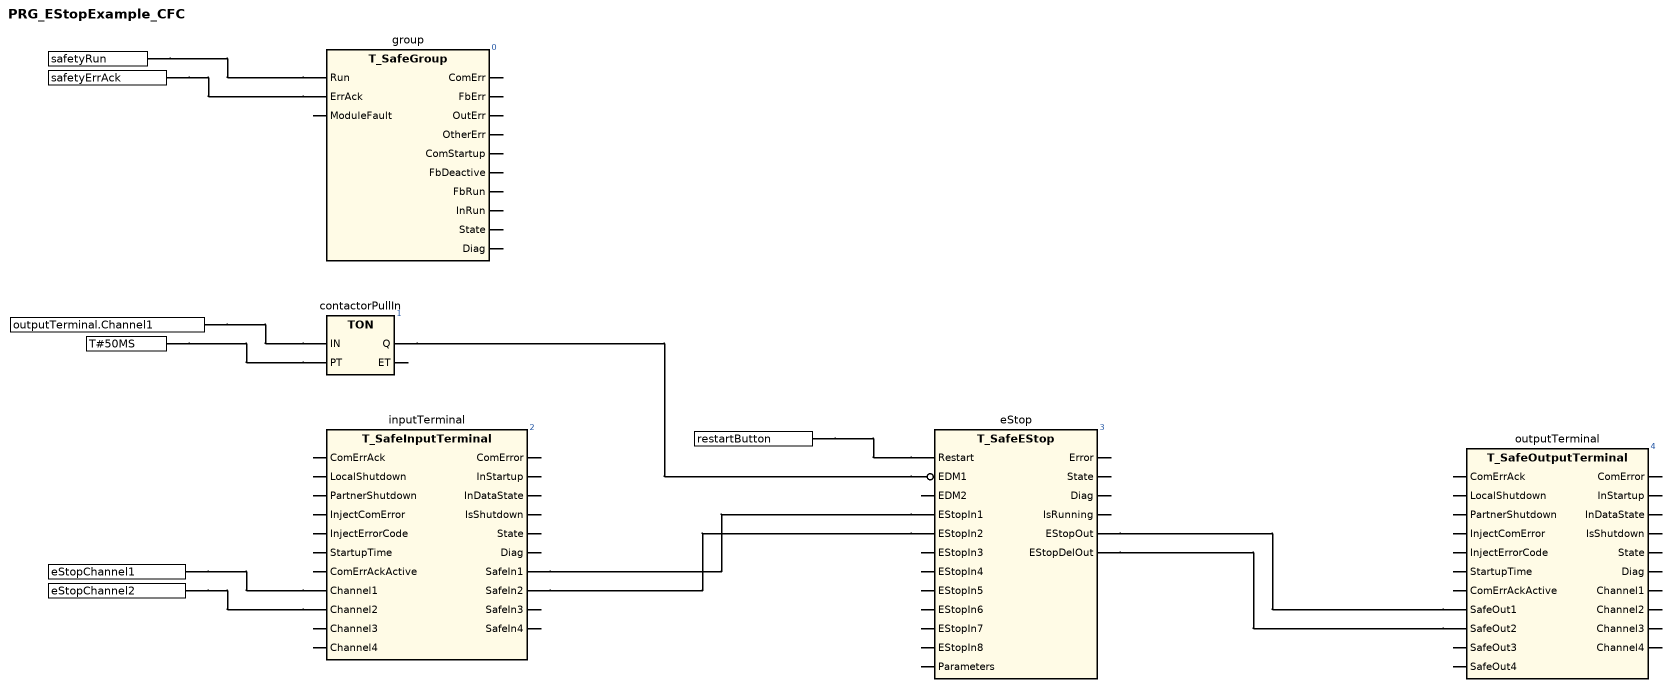
group(Run := safetyRun, ErrAck := safetyErrAck); // T_SafeGroup
contactorPullIn(IN := outputTerminal.Channel1, PT := T#50MS); // TON
inputTerminal(Channel1 := eStopChannel1, Channel2 := eStopChannel2); // T_SafeInputTerminal
eStop(
    Restart := restartButton,
    EDM1 := NOT contactorPullIn.Q,
    EStopIn1 := inputTerminal.SafeIn1,
    EStopIn2 := inputTerminal.SafeIn2); // T_SafeEStop
outputTerminal(SafeOut1 := eStop.EStopOut, SafeOut2 := eStop.EStopDelOut); // T_SafeOutputTerminal

END_PROGRAM

// FunctionBlocks/T_SafeConnShutdown
// Model of the TwinSAFE FB CONNECTION SHUTDOWN.
// Shuts down the assigned connection while the Deactivate inputs are TRUE and reports Deactivated
// once the connection is shut down (also when the partner shut it down). The connection is assigned
// at construction (the Connection ID of the Safety Editor):
//     connShutdown : T_SafeConnShutdown(group := safetyGroup, connection := toolConnection);
{attribute 'reflection'}
FUNCTION_BLOCK T_SafeConnShutdown EXTENDS T_SafeFunctionBlockBase
VAR_INPUT
    Deactivate1 : BOOL;
    Deactivate2 : BOOL;
    Parameters : ST_SafeConnShutdownParameters;
END_VAR
VAR_OUTPUT
    Deactivated : BOOL;
END_VAR
VAR
    {attribute 'is_connected' := 'Deactivate1'}
    _deactivate1Connected : BOOL;
    {attribute 'is_connected' := 'Deactivate2'}
    _deactivate2Connected : BOOL;
    _connection : REFERENCE TO T_SafeConnection;
    _pairs : ARRAY[1..1] OF T_SafeInputPair;
    _state : E_SafeFbState := E_SafeFbState.Stop;
    _prevState : E_SafeFbState;
END_VAR

SUPER^();

PROPERTY ConnShutdownState : E_SafeFbState
GET
ConnShutdownState := _state;
END_GET
END_PROPERTY

METHOD FB_init : BOOL
VAR_INPUT
    bInitRetains : BOOL;
    bInCopyCode : BOOL;
    group : REFERENCE TO T_SafeGroup; // the TwinSAFE group this block belongs to
    connection : REFERENCE TO T_SafeConnection; // the connection to shut down (Connection ID)
END_VAR
// the base FB_init (group registration) is called implicitly by TwinCAT
_connection REF= connection;
END_METHOD

METHOD PROTECTED Process
VAR
    acknowledge : BOOL;
    deactivate : BOOL;
    operating : BOOL;
    stateBefore : E_SafeFbState;
    passes : USINT;
END_VAR
acknowledge := (_state = E_SafeFbState.Error) AND _errAck;
_pairs[1](
    In1 := Deactivate1,
    In2 := Deactivate2,
    Active1 := _deactivate1Connected,
    Active2 := _deactivate2Connected,
    MakeContact1 := Parameters.Deactivate1MakeContact,
    MakeContact2 := Parameters.Deactivate2MakeContact,
    DiscrepancyTime := Parameters.DiscrepancyTime,
    Monitor := _fbRun,
    SafeInputsAfterDiscError := Parameters.SafeInputsAfterDiscError,
    Acknowledge := acknowledge
);

deactivate := _pairs[1].IsActive AND _pairs[1].AllTrue;

IF NOT _fbRun AND _state <> E_SafeFbState.Error AND _state <> E_SafeFbState.Reset THEN
    _state := E_SafeFbState.Stop;
END_IF

operating := (_state = E_SafeFbState.Safe) OR (_state = E_SafeFbState.Run);

IF _pairs[1].DiscrepancyError AND operating THEN
    UpdateDiscrepancyDiag();
    _state := E_SafeFbState.Error;
END_IF

passes := 0;

REPEAT
    stateBefore := _state;

    CASE _state OF
        E_SafeFbState.Stop:
            IF StateChanged() THEN
                Deactivated := FALSE;
                Error       := FALSE;
                Diag        := 0;
            END_IF

            _connection.LocalShutdown := FALSE;

            IF _fbRun THEN
                _state := E_SafeFbState.Safe;
            END_IF

        E_SafeFbState.Safe:
            IF StateChanged() THEN
                Deactivated := FALSE;
            END_IF

            _connection.LocalShutdown := deactivate;

            IF _connection.IsShutdown THEN
                _state := E_SafeFbState.Run;
            END_IF

        E_SafeFbState.Run:
            IF StateChanged() THEN
                Deactivated := TRUE;
            END_IF

            _connection.LocalShutdown := deactivate;

            IF NOT _connection.IsShutdown THEN
                _state := E_SafeFbState.Safe;
            END_IF

        E_SafeFbState.Error:
            IF StateChanged() THEN
                Deactivated := FALSE;
                Error       := TRUE;
            END_IF

            _connection.LocalShutdown := FALSE;
            UpdateDiscrepancyDiag();

            IF _errAck AND NOT _pairs[1].DiscrepancyError THEN
                _state := E_SafeFbState.Reset;
            END_IF

        E_SafeFbState.Reset:
            IF StateChanged() THEN
                Error := FALSE;
                Diag  := 0;
            END_IF

            IF _errAckFallingEdge THEN
                _state := SEL(_fbRun, E_SafeFbState.Stop, E_SafeFbState.Safe);
            END_IF
    END_CASE

    passes := passes + 1;
UNTIL (stateBefore = _state) OR (passes >= 3)
END_REPEAT

State := TO_BYTE(_state);
END_METHOD

METHOD PRIVATE StateChanged : BOOL
IF _prevState = _state THEN
    RETURN;
END_IF

_prevState   := _state;
StateChanged := TRUE;
END_METHOD

// Mirrors the discrepancy state of every pair into the diagnostic bits.
METHOD PRIVATE UpdateDiscrepancyDiag
VAR
    i : USINT;
END_VAR
FOR i := 1 TO 1 DO
    IF _pairs[i].DiscrepancyError THEN
        SetDiagBit(0);

        IF _pairs[i].AwaitingSafeInputs THEN
            SetDiagBit(8);
        ELSE
            ClearDiagBit(8);
        END_IF
    END_IF
END_FOR
END_METHOD

END_FUNCTION_BLOCK

// FunctionBlocks/T_SafeDecouple
// Model of the TwinSAFE FB DECOUPLE: eight inputs looped one-to-one to eight outputs.
FUNCTION_BLOCK T_SafeDecouple EXTENDS T_SafeFunctionBlockBase
VAR_INPUT
    DecIn1 : BOOL;
    DecIn2 : BOOL;
    DecIn3 : BOOL;
    DecIn4 : BOOL;
    DecIn5 : BOOL;
    DecIn6 : BOOL;
    DecIn7 : BOOL;
    DecIn8 : BOOL;
END_VAR
VAR_OUTPUT
    DecOut1 : BOOL;
    DecOut2 : BOOL;
    DecOut3 : BOOL;
    DecOut4 : BOOL;
    DecOut5 : BOOL;
    DecOut6 : BOOL;
    DecOut7 : BOOL;
    DecOut8 : BOOL;
END_VAR
VAR
    _state : E_SafeFbState := E_SafeFbState.Stop;
END_VAR

SUPER^();

METHOD PROTECTED Process
VAR
    run : BOOL;
END_VAR
run     := _fbRun;
_state  := SEL(run, E_SafeFbState.Stop, E_SafeFbState.Run);
DecOut1 := run AND DecIn1;
DecOut2 := run AND DecIn2;
DecOut3 := run AND DecIn3;
DecOut4 := run AND DecIn4;
DecOut5 := run AND DecIn5;
DecOut6 := run AND DecIn6;
DecOut7 := run AND DecIn7;
DecOut8 := run AND DecIn8;
Error   := FALSE;
Diag    := 0;
State   := TO_BYTE(_state);
END_METHOD

END_FUNCTION_BLOCK

// FunctionBlocks/T_SafeEdm
// Model of the TwinSAFE FB EDM (external device monitor):
// Mon2 must take the opposite value to Mon1 within the configured switch-on / switch-off time.
// The Safety Editor refuses an EDM with Mon1 or Mon2 unconnected: the model then reports Error with
// diagnostic bit 15 instead of running (see T_SafeFunctionBlockBase).
{attribute 'reflection'}
FUNCTION_BLOCK T_SafeEdm EXTENDS T_SafeFunctionBlockBase
VAR_INPUT
    Mon1 : BOOL;
    Mon2 : BOOL;
    Parameters : ST_SafeEdmParameters;
END_VAR
VAR
    {attribute 'is_connected' := 'Mon1'}
    _mon1Connected : BOOL;
    {attribute 'is_connected' := 'Mon2'}
    _mon2Connected : BOOL;
    _state : E_SafeEdmState := E_SafeEdmState.Stop;
    _prevState : E_SafeEdmState;
    _timer : TON;
    _satisfied : BOOL;
END_VAR

SUPER^();
IsRunning := (_state = E_SafeEdmState.MonOn) OR (_state = E_SafeEdmState.MonOff);

// Mon1 and Mon2 must both be connected (Safety Editor: "Inport Mon1 of EDM must be connected").
METHOD PROTECTED ConfigurationOk : BOOL
IF NOT _mon1Connected THEN
    _configurationFault := 'T_SafeEdm: Inport Mon1 of EDM must be connected';
    RETURN;
ELSIF NOT _mon2Connected THEN
    _configurationFault := 'T_SafeEdm: Inport Mon2 of EDM must be connected';
    RETURN;
END_IF

ConfigurationOk := TRUE;
END_METHOD

METHOD PROTECTED Process
VAR
    monitor1 : BOOL;
    monitor2 : BOOL;
    stateBefore : E_SafeEdmState;
    passes : USINT;
END_VAR
monitor1 := F_SafeInputValue(_mon1Connected, Parameters.Mon1MakeContact, Mon1);
monitor2 := F_SafeInputValue(_mon2Connected, Parameters.Mon2MakeContact, Mon2);

IF NOT _fbRun AND _state <> E_SafeEdmState.Error AND _state <> E_SafeEdmState.Reset THEN
    _state := E_SafeEdmState.Stop;
END_IF

passes := 0;

REPEAT
    stateBefore := _state;

    CASE _state OF
        E_SafeEdmState.Stop:
            IF StateChanged() THEN
                Error := FALSE;
                Diag  := 0;
                _timer(IN := FALSE, PT := T#0S);
            END_IF

            IF _fbRun THEN
                _state := SEL(monitor1, E_SafeEdmState.MonOff, E_SafeEdmState.MonOn);
            END_IF

        E_SafeEdmState.MonOn:
            // switch-on monitoring: Mon2 must become FALSE within SwitchOnTime
            IF StateChanged() THEN
                _satisfied := FALSE;
                _timer(IN := FALSE, PT := Parameters.SwitchOnTime);
            END_IF

            IF NOT monitor2 THEN
                _satisfied := TRUE;
            END_IF

            _timer(IN := NOT _satisfied AND (Parameters.SwitchOnTime > T#0S), PT := Parameters.SwitchOnTime);

            IF _timer.Q THEN
                SetDiagBit(1);
                _state := E_SafeEdmState.Error;
            ELSIF NOT monitor1 THEN
                _state := E_SafeEdmState.MonOff;
            END_IF

        E_SafeEdmState.MonOff:
            // switch-off monitoring: Mon2 must become TRUE within SwitchOffTime
            IF StateChanged() THEN
                _satisfied := FALSE;
                _timer(IN := FALSE, PT := Parameters.SwitchOffTime);
            END_IF

            IF monitor2 THEN
                _satisfied := TRUE;
            END_IF

            _timer(IN := NOT _satisfied AND (Parameters.SwitchOffTime > T#0S), PT := Parameters.SwitchOffTime);

            IF _timer.Q THEN
                SetDiagBit(0);
                _state := E_SafeEdmState.Error;
            ELSIF monitor1 THEN
                _state := E_SafeEdmState.MonOn;
            END_IF

        E_SafeEdmState.Error:
            IF StateChanged() THEN
                Error := TRUE;
                _timer(IN := FALSE, PT := T#0S);
            END_IF

            IF _errAck THEN
                _state := E_SafeEdmState.Reset;
            END_IF

        E_SafeEdmState.Reset:
            IF StateChanged() THEN
                Error := FALSE;
                Diag  := 0;
            END_IF

            IF _errAckFallingEdge THEN
                IF NOT _fbRun THEN
                    _state := E_SafeEdmState.Stop;
                ELSE
                    _state := SEL(monitor1, E_SafeEdmState.MonOff, E_SafeEdmState.MonOn);
                END_IF
            END_IF
    END_CASE

    passes := passes + 1;
UNTIL (stateBefore = _state) OR (passes >= 3)
END_REPEAT

State := TO_BYTE(_state);
END_METHOD

METHOD PRIVATE StateChanged : BOOL
IF _prevState = _state THEN
    RETURN;
END_IF

_prevState   := _state;
StateChanged := TRUE;
END_METHOD

END_FUNCTION_BLOCK

// FunctionBlocks/T_SafeMon
// Model of the TwinSAFE FB MON (safety door / guard monitoring).
// Two MonIn pairs, a Secure pair that bypasses them, manual restart (when Restart is connected),
// manual function test, two EDM feedback loops and a delayed output.
// The Safety Editor refuses a MON with no MonIn port connected, or an EDM reset time that is not 0 ms,
// a multiple of 10 ms and at most 60000 ms: the model then reports Error with diagnostic bit 15
// instead of running (see T_SafeFunctionBlockBase).
{attribute 'reflection'}
FUNCTION_BLOCK T_SafeMon EXTENDS T_SafeFunctionBlockBase
VAR_INPUT
    Restart : BOOL; // connect for manual restart; may be a standard PLC signal
    EDM1 : BOOL; // feedback loop of MonOut
    EDM2 : BOOL; // feedback loop of MonDelOut
    MonIn1 : BOOL;
    MonIn2 : BOOL;
    MonIn3 : BOOL;
    MonIn4 : BOOL;
    Secure1 : BOOL; // when TRUE (after normalisation) the MonIn inputs are ignored
    Secure2 : BOOL;
    Parameters : ST_SafeMonParameters;
END_VAR
VAR_OUTPUT
    MonOut : BOOL;
    MonDelOut : BOOL;
END_VAR
VAR
    {attribute 'is_connected' := 'Restart'}
    _restartConnected : BOOL;
    {attribute 'is_connected' := 'EDM1'}
    _eDM1Connected : BOOL;
    {attribute 'is_connected' := 'EDM2'}
    _eDM2Connected : BOOL;
    {attribute 'is_connected' := 'MonIn1'}
    _monIn1Connected : BOOL;
    {attribute 'is_connected' := 'MonIn2'}
    _monIn2Connected : BOOL;
    {attribute 'is_connected' := 'MonIn3'}
    _monIn3Connected : BOOL;
    {attribute 'is_connected' := 'MonIn4'}
    _monIn4Connected : BOOL;
    {attribute 'is_connected' := 'Secure1'}
    _secure1Connected : BOOL;
    {attribute 'is_connected' := 'Secure2'}
    _secure2Connected : BOOL;
    _pairs : ARRAY[1..3] OF T_SafeInputPair; // 1: MonIn1/2, 2: MonIn3/4, 3: Secure1/2
    _state : E_SafeMonState := E_SafeMonState.Stop;
    _prevState : E_SafeMonState;
    _restartPrev : BOOL;
    _delayTimer : TON;
    _delayRunning : BOOL;
    _funcTested : ARRAY[1..2] OF BOOL;
    _edmResetTimer1 : TON;
    _edmResetTimer2 : TON;
    _edm1Dropped : BOOL;
    _edm2Dropped : BOOL;
END_VAR

SUPER^();

// At least one MonIn port must be connected and the EDM reset times must be 0 ms or a multiple of 10 ms up to 60000 ms (Safety Editor messages).
METHOD PROTECTED ConfigurationOk : BOOL
IF NOT (_monIn1Connected OR _monIn2Connected OR _monIn3Connected OR _monIn4Connected) THEN
    _configurationFault := 'T_SafeMon: MON does not have at least 1 MonIn(x) port active and connected';
    RETURN;
ELSIF NOT F_SafeResetTimeOk(Parameters.Edm1ResetTime) THEN
    _configurationFault := 'T_SafeMon: $'Reset Time$' parameter of EDM1 of MON has to be 0 ms or a multiple of 10 ms and maximal 60000 ms';
    RETURN;
ELSIF NOT F_SafeResetTimeOk(Parameters.Edm2ResetTime) THEN
    _configurationFault := 'T_SafeMon: $'Reset Time$' parameter of EDM2 of MON has to be 0 ms or a multiple of 10 ms and maximal 60000 ms';
    RETURN;
END_IF

ConfigurationOk := TRUE;
END_METHOD

// Checks the EDM inputs at restart and records diagnostic bits 4/5 on failure.
METHOD PRIVATE EdmInputsOk : BOOL
EdmInputsOk := TRUE;

IF _eDM1Connected AND NOT EDM1 THEN
    SetDiagBit(4);
    EdmInputsOk := FALSE;
END_IF

IF _eDM2Connected AND NOT EDM2 THEN
    SetDiagBit(5);
    EdmInputsOk := FALSE;
END_IF
END_METHOD

// TRUE when every connected EDM input reads 1 (contactors released).
METHOD PRIVATE EdmInputsTrue : BOOL
EdmInputsTrue := (NOT _eDM1Connected OR EDM1) AND (NOT _eDM2Connected OR EDM2);
END_METHOD

// EL6910 extension: after the outputs switch on, each connected EDM input must drop to FALSE
// within its Reset Time. Returns FALSE (and sets diagnostic bits 4/5) on timeout.
METHOD PRIVATE EdmResetOk : BOOL
EdmResetOk := TRUE;

IF _eDM1Connected AND Parameters.Edm1ResetTime > T#0S THEN
    IF NOT EDM1 THEN
        _edm1Dropped := TRUE;
    END_IF

    _edmResetTimer1(IN := NOT _edm1Dropped, PT := Parameters.Edm1ResetTime);

    IF _edmResetTimer1.Q THEN
        SetDiagBit(4);
        EdmResetOk := FALSE;
    END_IF
END_IF

IF _eDM2Connected AND Parameters.Edm2ResetTime > T#0S THEN
    IF NOT EDM2 THEN
        _edm2Dropped := TRUE;
    END_IF

    _edmResetTimer2(IN := NOT _edm2Dropped, PT := Parameters.Edm2ResetTime);

    IF _edmResetTimer2.Q THEN
        SetDiagBit(5);
        EdmResetOk := FALSE;
    END_IF
END_IF
END_METHOD

PROPERTY MonState : E_SafeMonState
GET
MonState := _state;
END_GET
END_PROPERTY

METHOD PROTECTED Process
VAR
    i : USINT;
    acknowledge : BOOL;
    monRequested : BOOL;
    bypass : BOOL;
    safeRequested : BOOL;
    discError : BOOL;
    restartFalling : BOOL;
    functionTestDue : BOOL;
    stateBefore : E_SafeMonState;
    passes : USINT;
END_VAR
acknowledge := (_state = E_SafeMonState.Error) AND _errAck;
_pairs[1](
    In1 := MonIn1,
    In2 := MonIn2,
    Active1 := _monIn1Connected,
    Active2 := _monIn2Connected,
    MakeContact1 := Parameters.MonIn1MakeContact,
    MakeContact2 := Parameters.MonIn2MakeContact,
    DiscrepancyTime := Parameters.DiscrepancyTime1,
    Monitor := _fbRun,
    SafeInputsAfterDiscError := Parameters.SafeInputsAfterDiscError,
    Acknowledge := acknowledge
);

_pairs[2](
    In1 := MonIn3,
    In2 := MonIn4,
    Active1 := _monIn3Connected,
    Active2 := _monIn4Connected,
    MakeContact1 := Parameters.MonIn3MakeContact,
    MakeContact2 := Parameters.MonIn4MakeContact,
    DiscrepancyTime := Parameters.DiscrepancyTime2,
    Monitor := _fbRun,
    SafeInputsAfterDiscError := Parameters.SafeInputsAfterDiscError,
    Acknowledge := acknowledge
);

_pairs[3](
    In1 := Secure1,
    In2 := Secure2,
    Active1 := _secure1Connected,
    Active2 := _secure2Connected,
    MakeContact1 := Parameters.Secure1MakeContact,
    MakeContact2 := Parameters.Secure2MakeContact,
    DiscrepancyTime := Parameters.SecureDiscrepancyTime,
    Monitor := _fbRun,
    SafeInputsAfterDiscError := Parameters.SafeInputsAfterDiscError,
    Acknowledge := acknowledge
);

monRequested  := _pairs[1].SafeStateRequested OR _pairs[2].SafeStateRequested;
bypass        := _pairs[3].IsActive AND _pairs[3].AllTrue;
safeRequested := monRequested AND NOT bypass;

FOR i := 1 TO 3 DO
    discError := discError OR _pairs[i].DiscrepancyError;
END_FOR

restartFalling := NOT Restart AND _restartPrev;
_restartPrev   := Restart;

IF NOT _fbRun AND _state <> E_SafeMonState.Error AND _state <> E_SafeMonState.Reset THEN
    _state := E_SafeMonState.Stop;
END_IF

// Discrepancy errors: immediate, except that a running delayed output completes its delay first
IF discError THEN
    CASE _state OF
        E_SafeMonState.Safe, E_SafeMonState.Start, E_SafeMonState.FuncTest:
            UpdateDiscrepancyDiag();
            _state := E_SafeMonState.Error;
        E_SafeMonState.Run:
            UpdateDiscrepancyDiag();

            IF Parameters.DelayTime > T#0S THEN
                _state := E_SafeMonState.ErrorDelay;
            ELSE
                _state := E_SafeMonState.Error;
            END_IF
        E_SafeMonState.DelayOut:
            UpdateDiscrepancyDiag();
            _state := E_SafeMonState.ErrorDelay;
    END_CASE
END_IF

passes := 0;

REPEAT
    stateBefore := _state;

    CASE _state OF
        E_SafeMonState.Stop:
            IF StateChanged() THEN
                SetOutputsSafe();
                Error          := FALSE;
                Diag           := 0;
                _delayRunning  := FALSE;
                _funcTested[1] := FALSE;
                _funcTested[2] := FALSE;
            END_IF

            IF _fbRun THEN
                functionTestDue := Parameters.ManualFunctionTest AND (_pairs[1].IsActive OR _pairs[2].IsActive);
                _state          := SEL(functionTestDue, E_SafeMonState.Safe, E_SafeMonState.FuncTest);
            END_IF

        E_SafeMonState.FuncTest:
            // every connected MonIn pair must request the safe state once before a restart is accepted
            IF StateChanged() THEN
                SetOutputsSafe();
            END_IF

            IF _pairs[1].SafeStateRequested THEN
                _funcTested[1] := TRUE;
            END_IF

            IF _pairs[2].SafeStateRequested THEN
                _funcTested[2] := TRUE;
            END_IF

            IF (NOT _pairs[1].IsActive OR _funcTested[1]) AND (NOT _pairs[2].IsActive OR _funcTested[2]) THEN
                _state := E_SafeMonState.Safe;
            END_IF

        E_SafeMonState.Safe:
            IF StateChanged() THEN
                SetOutputsSafe();
                _delayRunning := FALSE;
            END_IF

            IF _restartConnected THEN
                IF Restart THEN
                    IF NOT EdmInputsOk() THEN
                        _state := E_SafeMonState.Error;
                    ELSIF NOT safeRequested THEN
                        _state := E_SafeMonState.Start;
                    END_IF
                END_IF
            ELSIF NOT safeRequested AND EdmInputsTrue() THEN
                // automatic restart: an EDM fault keeps the FB in SAFE without an error
                _state := E_SafeMonState.Run;
            END_IF

        E_SafeMonState.Start:
            IF StateChanged() THEN
                SetOutputsSafe();
            END_IF

            IF safeRequested THEN
                _state := E_SafeMonState.Safe;
            ELSIF restartFalling THEN
                IF EdmInputsOk() THEN
                    _state := E_SafeMonState.Run;
                ELSE
                    _state := E_SafeMonState.Error;
                END_IF
            END_IF

        E_SafeMonState.Run:
            IF StateChanged() THEN
                MonOut    := TRUE;
                MonDelOut := TRUE;
                StartEdmResetMonitoring();
            END_IF

            IF NOT EdmResetOk() THEN
                _state := E_SafeMonState.Error;
            ELSIF safeRequested THEN
                IF Parameters.DelayTime > T#0S THEN
                    _state := E_SafeMonState.DelayOut;
                ELSE
                    _state := E_SafeMonState.Safe;
                END_IF
            END_IF

        E_SafeMonState.DelayOut:
            IF StateChanged() THEN
                MonOut    := FALSE;
                MonDelOut := TRUE;
                _delayTimer(IN := FALSE, PT := Parameters.DelayTime);
                _delayRunning := TRUE;
            END_IF

            _delayTimer(IN := TRUE, PT := Parameters.DelayTime);

            IF _delayTimer.Q THEN
                _state := E_SafeMonState.Safe;
            END_IF

        E_SafeMonState.ErrorDelay:
            IF StateChanged() THEN
                MonOut    := FALSE;
                MonDelOut := TRUE;

                IF NOT _delayRunning THEN
                    _delayTimer(IN := FALSE, PT := Parameters.DelayTime);
                    _delayRunning := TRUE;
                END_IF
            END_IF

            _delayTimer(IN := TRUE, PT := Parameters.DelayTime);

            IF _delayTimer.Q THEN
                _state := E_SafeMonState.Error;
            END_IF

        E_SafeMonState.Error:
            IF StateChanged() THEN
                SetOutputsSafe();
                Error         := TRUE;
                _delayRunning := FALSE;
            END_IF

            UpdateDiscrepancyDiag();

            IF _errAck AND NOT discError THEN
                _state := E_SafeMonState.Reset;
            END_IF

        E_SafeMonState.Reset:
            IF StateChanged() THEN
                SetOutputsSafe();
                Error := FALSE;
                Diag  := 0;
            END_IF

            IF _errAckFallingEdge THEN
                _state := SEL(_fbRun, E_SafeMonState.Stop, E_SafeMonState.Safe);
            END_IF
    END_CASE

    passes := passes + 1;
UNTIL (stateBefore = _state) OR (passes >= 3)
END_REPEAT

State := TO_BYTE(_state);
END_METHOD

METHOD PRIVATE SetOutputsSafe
MonOut    := FALSE;
MonDelOut := FALSE;
END_METHOD

METHOD PRIVATE StartEdmResetMonitoring
_edm1Dropped := FALSE;
_edm2Dropped := FALSE;
_edmResetTimer1(IN := FALSE, PT := Parameters.Edm1ResetTime);
_edmResetTimer2(IN := FALSE, PT := Parameters.Edm2ResetTime);
END_METHOD

METHOD PRIVATE StateChanged : BOOL
IF _prevState = _state THEN
    RETURN;
END_IF

_prevState   := _state;
StateChanged := TRUE;
END_METHOD

// Mirrors the discrepancy state of every pair into the diagnostic bits.
METHOD PRIVATE UpdateDiscrepancyDiag
VAR
    i : USINT;
END_VAR
FOR i := 1 TO 3 DO
    IF _pairs[i].DiscrepancyError THEN
        SetDiagBit(i - 1);

        IF _pairs[i].AwaitingSafeInputs THEN
            SetDiagBit(i + 7);
        ELSE
            ClearDiagBit(i + 7);
        END_IF
    END_IF
END_FOR
END_METHOD

END_FUNCTION_BLOCK

